(* IEC 61131-3 sources: TetherPLC/compat/tc3 (part 3) *)

(* ---- tc3_mc2_ah.st ---- *)
// Tc3_MC2_AdvancedHoming — user-programmable homing sequences.
//
// All 16 documented APIs over the builtin FB_MotionAxis
// (tplc-motion service), flattened to this dialect:
//
//   AXIS_REF                -> Axis : UDINT (FB_MotionAxis handle)
//   MC_HomingParameter      -> 15 VAR_IN_OUT members P_* (Stored flag
//                             plus the NC soft-limit/lag/vel-diff and
//                             drive torque Stored/Actual fields; the
//                             sim exposes no such drive params so the
//                             fields are pass-through bookkeeping)
//   MC_Ref_Signal_Ref       -> RefLevel : BOOL (the .Level member;
//                             SignalSource/TouchProbe have no sim
//                             equivalent and are dropped)
//   MC_Home_Direction       -> Direction : UDINT
//                             (1=mcPositiveDirection, 3=mcNegative-
//                             Direction, 5=mcSwitchPositive,
//                             7=mcSwitchNegative)
//   MC_Switch_Mode          -> SwitchMode : UDINT
//                             (1=mcOn, 2=mcOff, 3=mcRisingEdge,
//                             4=mcFallingEdge, 5=mcEdgeSwitchPositive,
//                             6=mcEdgeSwitchNegative,
//                             11=mcRisingEdgeInverse,
//                             12=mcFallingEdgeInverse)
//   MC_BufferMode           -> BufferMode : UDINT (not implemented,
//                             accepted and ignored like TwinCAT)
//   ST_Home_Options         -> (empty struct, no member)
//   ST_Home_Options2        -> OptDisableDriveAccess : BOOL
//   ST_Home_Options3        -> OptDisableDriveAccess +
//                             OptInstantLagReduction : BOOL
//   ST_Home_Options4        -> OptDisableDriveAccess +
//                             OptEnableLagErrorDetection : BOOL
//   E_HomingErrorCodes      -> ErrorID values 16#4B90..16#4B98
//
// Motion model: step FBs run a PV-mode (0x6060=3) velocity search at
// Velocity user units/s (0x60FF), poll the OP6 snapshot, and evaluate
// the switch/block condition each scan.  On detection the axis is
// stopped (0x60FF=0), allowed to settle, then the position is assigned
// via a direct 0x6064 write (MC_SetPosition equivalent) unless the FB
// is a "..Detection" variant, which instead returns RecordedPosition.
// The sensor "signal" is the user-fed RefLevel BOOL; the sim has no
// physical switch/encoder inputs.  Block detection uses the
// velocity-undershoot criterion (|VEL_ACTUAL| below
// DetectionVelocityLimit for DetectionVelocityTime); the travel-limit
// clamp added to the velocity modes makes a fixed stop produce that
// undershoot.  TorqueLimit/LagLimit/Acceleration/Deceleration/Jerk are
// accepted but inert (no torque or jerk model in the sim; PV ramps at
// the axis' configured accel/decel).
//
// Internal engine: AH_Run.  Kind codes: 1 absSwitch, 2 absSwitchDet,
// 3 block, 4 blockDet, 5 blockLag, 6 blockLagDet, 7 limitSwitch,
// 8 limitSwitchDet, 9 refPulse, 10 refPulseDet, 11 flyingRefPulse,
// 12 flyingSwitch, 20 distance move (FinishHoming).

// ---- AH_Run: shared homing sequence engine (internal helper) ----
FUNCTION_BLOCK AH_Run
VAR_INPUT
    Execute : BOOL;
    Axis : UDINT;
    Kind : UDINT;
    Direction : UDINT;
    SwitchMode : UDINT;
    RefLevel : BOOL;
    Velocity : LREAL;
    SetPosEn : BOOL;
    SetPosition : LREAL;
    TimeLimit : TIME;
    DistanceLimit : LREAL;
    DetVelLimit : LREAL;
    DetVelTime : TIME;
    LagLimit : LREAL;
    PosLimSw : BOOL;
    NegLimSw : BOOL;
    Distance : LREAL;
    ParamIn : BOOL;
END_VAR
VAR_OUTPUT
    Done : BOOL;
    Busy : BOOL;
    Active : BOOL;
    CommandAborted : BOOL;
    Error : BOOL;
    ErrorID : UDINT;
    RecordedPosition : LREAL;
    ParamOut : BOOL;
END_VAR
VAR
    ax : FB_MotionAxis;
    clk : TON;
    exPrev : BOOL;
    phase : UDINT;          // 0 idle, 1 search, 2 settle, 3 distmove, 4 observe
    refPrev : BOOL;
    moveDir : DINT;
    startPos : DINT;
    startNs : LINT;
    detNs : LINT;           // undershoot start, -1 = not undershooting
    velCmd : DINT;
    pendSet : BOOL;
    recPos : LREAL;
    distGoal : DINT;
    nowNs : LINT;
    pos : DINT;
    vel : DINT;
    cond : BOOL;
    isSwitch : BOOL;
    isBlock : BOOL;
    isDet : BOOL;
    edge : BOOL;
    pStored : BOOL;
END_VAR
    clk(IN := TRUE, PT := T#1000000h);
    ax.AXIS := Axis;
    ax.OP := 3; ax();
    ax.OP := 6; ax();
    Done := FALSE; Busy := FALSE; Active := FALSE;
    CommandAborted := FALSE; Error := FALSE; ErrorID := 0;
    RecordedPosition := 0.0;
    nowNs := TIME_TO_LINT(clk.ET);
    pos := ax.POS_ACTUAL;
    vel := ax.VEL_ACTUAL;
    pStored := ParamIn;
    isSwitch := (Kind >= 1) AND (Kind <= 2) OR (Kind >= 7) AND (Kind <= 10);
    isBlock := (Kind >= 3) AND (Kind <= 6);
    isDet := (Kind = 2) OR (Kind = 4) OR (Kind = 6) OR (Kind = 8)
             OR (Kind = 10);
    edge := Execute AND NOT exPrev;
    exPrev := Execute;

    IF phase = 0 THEN
        IF edge THEN
            // ---- validation ----
            IF Kind <> 11 AND Kind <> 12 AND Velocity <= 0.0 THEN
                Error := TRUE; ErrorID := 16#4B93;   // MC_HOMINGERROR_MODE
            ELSIF Kind <= 12 AND DistanceLimit < 0.0 THEN
                Error := TRUE; ErrorID := 16#4B96;   // DISTANCELIMIT
            ELSIF (Kind >= 1) AND (Kind <= 10)
                  AND Direction <> 1 AND Direction <> 3
                  AND Direction <> 5 AND Direction <> 7 THEN
                Error := TRUE; ErrorID := 16#4B91;   // DIRECTION
            ELSIF isSwitch AND SwitchMode <> 1 AND SwitchMode <> 2
                  AND SwitchMode <> 3 AND SwitchMode <> 4
                  AND SwitchMode <> 5 AND SwitchMode <> 6
                  AND SwitchMode <> 11 AND SwitchMode <> 12 THEN
                Error := TRUE; ErrorID := 16#4B92;   // SWITCHMODE
            ELSE
                // ---- initialise sequence ----
                IF Kind = 20 THEN
                    // distance move (FinishHoming backoff)
                    IF Distance = 0.0 THEN
                        pStored := FALSE;
                        Done := TRUE;
                    ELSE
                        moveDir := 1;
                        IF Distance < 0.0 THEN moveDir := -1; END_IF;
                        startPos := pos; startNs := nowNs; detNs := -1;
                        distGoal := pos + LREAL_TO_DINT(Distance);
                        refPrev := RefLevel;
                        pStored := TRUE;
                        velCmd := LREAL_TO_DINT(DINT_TO_LREAL(moveDir)
                                                * Velocity);
                        ax.OP := 5; ax.INDEX := 16#6060; ax.VALUE := 3; ax();
                        ax.OP := 5; ax.INDEX := 16#60FF;
                        ax.VALUE := velCmd; ax();
                        ax.OP := 5; ax.INDEX := 16#6040;
                        ax.VALUE := 16#000F; ax();
                        IF ax.STATUS = 0 THEN
                            phase := 3; Active := TRUE;
                        ELSE
                            Error := TRUE; ErrorID := ax.ERRID;
                            pStored := FALSE;
                        END_IF;
                    END_IF;
                ELSIF Kind = 11 OR Kind = 12 THEN
                    // passive observation, no motion commanded
                    startPos := pos; startNs := nowNs; detNs := -1;
                    refPrev := RefLevel;
                    pStored := TRUE;
                    phase := 4; Active := TRUE;
                ELSE
                    // search move direction
                    moveDir := 1;
                    IF Direction = 3 THEN moveDir := -1; END_IF;
                    IF Direction = 5 THEN
                        moveDir := 1;
                        IF RefLevel THEN moveDir := -1; END_IF;
                    END_IF;
                    IF Direction = 7 THEN
                        moveDir := -1;
                        IF RefLevel THEN moveDir := 1; END_IF;
                    END_IF;
                    startPos := pos; startNs := nowNs; detNs := -1;
                    refPrev := RefLevel;
                    pStored := TRUE;
                    velCmd := LREAL_TO_DINT(DINT_TO_LREAL(moveDir)
                                            * Velocity);
                    ax.OP := 5; ax.INDEX := 16#6060; ax.VALUE := 3; ax();
                    ax.OP := 5; ax.INDEX := 16#60FF; ax.VALUE := velCmd; ax();
                    ax.OP := 5; ax.INDEX := 16#6040; ax.VALUE := 16#000F; ax();
                    IF ax.STATUS = 0 THEN
                        phase := 1; Active := TRUE;
                    ELSE
                        Error := TRUE; ErrorID := ax.ERRID;
                        pStored := FALSE;
                    END_IF;
                END_IF;
            END_IF;
        END_IF;

    ELSIF phase = 1 THEN
        // ---- search: abort limits then detection ----
        IF (TimeLimit > T#0s) AND
           (nowNs - startNs > TIME_TO_LINT(TimeLimit)) THEN
            ax.OP := 5; ax.INDEX := 16#60FF; ax.VALUE := 0; ax();
            phase := 0; CommandAborted := TRUE;
        ELSIF ABS(DINT_TO_LREAL(pos - startPos)) > DistanceLimit THEN
            ax.OP := 5; ax.INDEX := 16#60FF; ax.VALUE := 0; ax();
            phase := 0; CommandAborted := TRUE;
        ELSIF (PosLimSw AND moveDir > 0) OR (NegLimSw AND moveDir < 0) THEN
            ax.OP := 5; ax.INDEX := 16#60FF; ax.VALUE := 0; ax();
            phase := 0; CommandAborted := TRUE;
        ELSE
            cond := FALSE;
            IF isSwitch THEN
                // MC_Switch_Mode evaluation; inverse variants share
                // the physical edge (approach side is absorbed by
                // the position assignment)
                IF SwitchMode = 1 THEN
                    cond := RefLevel;
                ELSIF SwitchMode = 2 THEN
                    cond := NOT RefLevel;
                ELSIF SwitchMode = 3 OR SwitchMode = 11 THEN
                    cond := RefLevel AND NOT refPrev;
                ELSIF SwitchMode = 4 OR SwitchMode = 12 THEN
                    cond := NOT RefLevel AND refPrev;
                ELSIF SwitchMode = 5 THEN
                    IF moveDir > 0 THEN
                        cond := RefLevel AND NOT refPrev;
                    ELSE
                        cond := NOT RefLevel AND refPrev;
                    END_IF;
                ELSIF SwitchMode = 6 THEN
                    IF moveDir > 0 THEN
                        cond := NOT RefLevel AND refPrev;
                    ELSE
                        cond := RefLevel AND NOT refPrev;
                    END_IF;
                END_IF;
            ELSIF isBlock THEN
                // velocity undershoot below DetVelLimit sustained
                // for DetVelTime; lag-based additionally requires
                // the velocity deficit proxy above LagLimit
                IF ABS(vel) < LREAL_TO_DINT(DetVelLimit) THEN
                    IF detNs < 0 THEN detNs := nowNs; END_IF;
                    IF nowNs - detNs >= TIME_TO_LINT(DetVelTime)
                       AND (Kind < 5 OR
                            ABS(velCmd - vel) > LREAL_TO_DINT(LagLimit)) THEN
                        cond := TRUE;
                    END_IF;
                ELSE
                    detNs := -1;
                END_IF;
            END_IF;
            refPrev := RefLevel;
            IF cond THEN
                ax.OP := 5; ax.INDEX := 16#60FF; ax.VALUE := 0; ax();
                recPos := DINT_TO_LREAL(pos);
                pendSet := SetPosEn AND NOT isDet;
                phase := 2; Active := TRUE;
            ELSE
                Active := TRUE; Busy := TRUE;
            END_IF;
        END_IF;

    ELSIF phase = 2 THEN
        // ---- settle: wait for the velocity ramp-down, then assign
        // the position (or report RecordedPosition) ----
        Active := TRUE; Busy := TRUE;
        IF ABS(vel) <= 1 THEN
            IF pendSet THEN
                ax.OP := 5; ax.INDEX := 16#6064;
                ax.VALUE := LREAL_TO_DINT(SetPosition); ax();
                IF ax.STATUS <> 0 THEN
                    Error := TRUE; ErrorID := ax.ERRID;
                    phase := 0;
                ELSE
                    phase := 0; Done := TRUE;
                    IF Kind = 20 THEN pStored := FALSE; END_IF;
                END_IF;
            ELSE
                IF isDet THEN RecordedPosition := recPos; END_IF;
                phase := 0; Done := TRUE;
                IF Kind = 20 THEN pStored := FALSE; END_IF;
            END_IF;
        END_IF;

    ELSIF phase = 3 THEN
        // ---- distance move: stop at the goal ----
        Active := TRUE; Busy := TRUE;
        IF (moveDir > 0 AND pos >= distGoal)
           OR (moveDir < 0 AND pos <= distGoal) THEN
            ax.OP := 5; ax.INDEX := 16#60FF; ax.VALUE := 0; ax();
            phase := 2;   // reuse settle; pendSet stays FALSE
            pendSet := FALSE;
        END_IF;
        IF (TimeLimit > T#0s) AND
           (nowNs - startNs > TIME_TO_LINT(TimeLimit)) THEN
            ax.OP := 5; ax.INDEX := 16#60FF; ax.VALUE := 0; ax();
            phase := 0; CommandAborted := TRUE; pStored := FALSE;
        END_IF;

    ELSIF phase = 4 THEN
        // ---- passive observation: no motion commanded ----
        Active := TRUE; Busy := TRUE;
        cond := FALSE;
        IF Kind = 11 THEN
            cond := RefLevel AND NOT refPrev;   // encoder zero pulse
        ELSE
            // flying switch: same MC_Switch_Mode evaluation,
            // direction taken as +1 (no search direction)
            IF SwitchMode = 1 THEN cond := RefLevel;
            ELSIF SwitchMode = 2 THEN cond := NOT RefLevel;
            ELSIF SwitchMode = 3 OR SwitchMode = 11 THEN
                cond := RefLevel AND NOT refPrev;
            ELSIF SwitchMode = 4 OR SwitchMode = 12 THEN
                cond := NOT RefLevel AND refPrev;
            ELSIF SwitchMode = 5 THEN
                cond := RefLevel AND NOT refPrev;
            ELSIF SwitchMode = 6 THEN
                cond := NOT RefLevel AND refPrev;
            END_IF;
        END_IF;
        refPrev := RefLevel;
        IF (TimeLimit > T#0s) AND
           (nowNs - startNs > TIME_TO_LINT(TimeLimit)) THEN
            phase := 0; CommandAborted := TRUE; pStored := FALSE;
        ELSIF ABS(DINT_TO_LREAL(pos - startPos)) > DistanceLimit THEN
            phase := 0; CommandAborted := TRUE; pStored := FALSE;
        ELSIF cond THEN
            ax.OP := 5; ax.INDEX := 16#6064;
            ax.VALUE := LREAL_TO_DINT(SetPosition); ax();
            IF ax.STATUS = 0 THEN
                phase := 0; Done := TRUE; pStored := FALSE;
            ELSE
                phase := 0; Error := TRUE; ErrorID := ax.ERRID;
                pStored := FALSE;
            END_IF;
        END_IF;
    END_IF;
    ParamOut := pStored;
END_FUNCTION_BLOCK

// ======================= finalizing FBs =======================

// MC_FinishHoming — completes a homing sequence: optional Distance
// backoff move at Velocity, then restores the stored parameters.
FUNCTION_BLOCK MC_FinishHoming
VAR_INPUT
    Execute : BOOL;
    Distance : LREAL;
    Velocity : LREAL;
    Acceleration : LREAL;
    Deceleration : LREAL;
    Jerk : LREAL;
    BufferMode : UDINT;
    OptDisableDriveAccess : BOOL;
END_VAR
VAR_IN_OUT
    Axis : UDINT;
    P_Stored : BOOL;
    P_NcSMin : BOOL;  P_NcSMax : BOOL;
    P_NcSPosDiff : BOOL;  P_NcSVeloDiff : BOOL;
    P_NcAMin : BOOL;  P_NcAMax : BOOL;
    P_NcAPosDiff : BOOL;  P_NcAVeloDiff : BOOL;
    P_DrvSBip : LREAL;  P_DrvSPos : LREAL;  P_DrvSNeg : LREAL;
    P_DrvABip : LREAL;  P_DrvAPos : LREAL;  P_DrvANeg : LREAL;
END_VAR
VAR_OUTPUT
    Done : BOOL;
    Busy : BOOL;
    CommandAborted : BOOL;
    Error : BOOL;
    ErrorID : UDINT;
END_VAR
VAR
    eng : AH_Run;
END_VAR
    eng.Execute := Execute; eng.Axis := Axis; eng.Kind := 20;
    eng.Direction := 1; eng.SwitchMode := 0; eng.RefLevel := FALSE;
    eng.Velocity := Velocity; eng.SetPosEn := FALSE;
    eng.SetPosition := 0.0;
    eng.TimeLimit := T#0s; eng.DistanceLimit := -1.0;
    eng.DetVelLimit := 0.0; eng.DetVelTime := T#0s; eng.LagLimit := 0.0;
    eng.PosLimSw := FALSE; eng.NegLimSw := FALSE;
    eng.Distance := Distance;
    eng.ParamIn := P_Stored;
    eng();
    P_Stored := eng.ParamOut;
    Done := eng.Done; Busy := eng.Busy;
    CommandAborted := eng.CommandAborted;
    Error := eng.Error; ErrorID := eng.ErrorID;
END_FUNCTION_BLOCK

// MC_HomeDirect — completes homing and assigns the axis position
// directly (no motion).  Axis leaves the homing state.
FUNCTION_BLOCK MC_HomeDirect
VAR_INPUT
    Execute : BOOL;
    SetPosition : LREAL;
    BufferMode : UDINT;
    OptDisableDriveAccess : BOOL;
END_VAR
VAR_IN_OUT
    Axis : UDINT;
    P_Stored : BOOL;
    P_NcSMin : BOOL;  P_NcSMax : BOOL;
    P_NcSPosDiff : BOOL;  P_NcSVeloDiff : BOOL;
    P_NcAMin : BOOL;  P_NcAMax : BOOL;
    P_NcAPosDiff : BOOL;  P_NcAVeloDiff : BOOL;
    P_DrvSBip : LREAL;  P_DrvSPos : LREAL;  P_DrvSNeg : LREAL;
    P_DrvABip : LREAL;  P_DrvAPos : LREAL;  P_DrvANeg : LREAL;
END_VAR
VAR_OUTPUT
    Done : BOOL;
    Busy : BOOL;
    Active : BOOL;
    CommandAborted : BOOL;
    Error : BOOL;
    ErrorID : UDINT;
END_VAR
VAR
    ax : FB_MotionAxis;
    exPrev : BOOL;
END_VAR
    ax.AXIS := Axis;
    Done := FALSE; Busy := FALSE; Active := FALSE;
    CommandAborted := FALSE; Error := FALSE; ErrorID := 0;
    IF Execute AND NOT exPrev THEN
        Active := TRUE;
        ax.OP := 5; ax.INDEX := 16#6064;
        ax.VALUE := LREAL_TO_DINT(SetPosition); ax();
        IF ax.STATUS = 0 THEN
            Done := TRUE; Active := FALSE;
            P_Stored := FALSE;
        ELSE
            Error := TRUE; ErrorID := ax.ERRID;
        END_IF;
    END_IF;
    exPrev := Execute;
END_FUNCTION_BLOCK

// MC_AbortHoming — aborts a homing sequence, stops any search move
// and restores the stored parameters.
FUNCTION_BLOCK MC_AbortHoming
VAR_INPUT
    Execute : BOOL;
    OptDisableDriveAccess : BOOL;
END_VAR
VAR_IN_OUT
    Axis : UDINT;
    P_Stored : BOOL;
    P_NcSMin : BOOL;  P_NcSMax : BOOL;
    P_NcSPosDiff : BOOL;  P_NcSVeloDiff : BOOL;
    P_NcAMin : BOOL;  P_NcAMax : BOOL;
    P_NcAPosDiff : BOOL;  P_NcAVeloDiff : BOOL;
    P_DrvSBip : LREAL;  P_DrvSPos : LREAL;  P_DrvSNeg : LREAL;
    P_DrvABip : LREAL;  P_DrvAPos : LREAL;  P_DrvANeg : LREAL;
END_VAR
VAR_OUTPUT
    Done : BOOL;
    Busy : BOOL;
    CommandAborted : BOOL;
    Error : BOOL;
    ErrorID : UDINT;
END_VAR
VAR
    ax : FB_MotionAxis;
    exPrev : BOOL;
END_VAR
    ax.AXIS := Axis;
    Done := FALSE; Busy := FALSE;
    CommandAborted := FALSE; Error := FALSE; ErrorID := 0;
    IF Execute AND NOT exPrev THEN
        ax.OP := 5; ax.INDEX := 16#60FF; ax.VALUE := 0; ax();
        ax.OP := 5; ax.INDEX := 16#6060; ax.VALUE := 0; ax();
        P_Stored := FALSE;
        Done := (ax.STATUS = 0);
        IF ax.STATUS <> 0 THEN Error := TRUE; ErrorID := ax.ERRID; END_IF;
    END_IF;
    exPrev := Execute;
END_FUNCTION_BLOCK

// ==================== referencing (passive) FBs ====================

// MC_AbortPassiveHoming — aborts passive homing.  The sim keeps no
// NC-side passive state, so this reports Done immediately.
FUNCTION_BLOCK MC_AbortPassiveHoming
VAR_INPUT
    Execute : BOOL;
END_VAR
VAR_IN_OUT
    Axis : UDINT;
END_VAR
VAR_OUTPUT
    Done : BOOL;
    Busy : BOOL;
    Active : BOOL;
    CommandAborted : BOOL;
    Error : BOOL;
    ErrorID : UDINT;
END_VAR
VAR
    exPrev : BOOL;
END_VAR
    Done := FALSE; Busy := FALSE; Active := FALSE;
    CommandAborted := FALSE; Error := FALSE; ErrorID := 0;
    IF Execute AND NOT exPrev THEN
        Done := TRUE;
    END_IF;
    exPrev := Execute;
END_FUNCTION_BLOCK

// MC_StepReferenceFlyingRefPulse — latch the position when the
// encoder zero pulse (RefLevel rising edge) arrives during an
// externally driven move, then assign SetPosition.
FUNCTION_BLOCK MC_StepReferenceFlyingRefPulse
VAR_INPUT
    Execute : BOOL;
    RefLevel : BOOL;
    SetPosition : LREAL;
    TimeLimit : TIME;
    DistanceLimit : LREAL;
    BufferMode : UDINT;
END_VAR
VAR_IN_OUT
    Axis : UDINT;
END_VAR
VAR_OUTPUT
    Done : BOOL;
    Busy : BOOL;
    Active : BOOL;
    CommandAborted : BOOL;
    Error : BOOL;
    ErrorID : UDINT;
END_VAR
VAR
    eng : AH_Run;
END_VAR
    eng.Execute := Execute; eng.Axis := Axis; eng.Kind := 11;
    eng.Direction := 1; eng.SwitchMode := 0; eng.RefLevel := RefLevel;
    eng.Velocity := 0.0; eng.SetPosEn := TRUE;
    eng.SetPosition := SetPosition;
    eng.TimeLimit := TimeLimit; eng.DistanceLimit := DistanceLimit;
    eng.DetVelLimit := 0.0; eng.DetVelTime := T#0s; eng.LagLimit := 0.0;
    eng.PosLimSw := FALSE; eng.NegLimSw := FALSE; eng.Distance := 0.0;
    eng.ParamIn := FALSE;
    eng();
    Done := eng.Done; Busy := eng.Busy; Active := eng.Active;
    CommandAborted := eng.CommandAborted;
    Error := eng.Error; ErrorID := eng.ErrorID;
END_FUNCTION_BLOCK

// MC_StepReferenceFlyingSwitch — same as FlyingRefPulse but the
// trigger is a MC_Switch_Mode condition on RefLevel.
FUNCTION_BLOCK MC_StepReferenceFlyingSwitch
VAR_INPUT
    Execute : BOOL;
    SwitchMode : UDINT;
    RefLevel : BOOL;
    SetPosition : LREAL;
    TimeLimit : TIME;
    DistanceLimit : LREAL;
    BufferMode : UDINT;
END_VAR
VAR_IN_OUT
    Axis : UDINT;
END_VAR
VAR_OUTPUT
    Done : BOOL;
    Busy : BOOL;
    Active : BOOL;
    CommandAborted : BOOL;
    Error : BOOL;
    ErrorID : UDINT;
END_VAR
VAR
    eng : AH_Run;
END_VAR
    eng.Execute := Execute; eng.Axis := Axis; eng.Kind := 12;
    eng.Direction := 1; eng.SwitchMode := SwitchMode;
    eng.RefLevel := RefLevel;
    eng.Velocity := 0.0; eng.SetPosEn := TRUE;
    eng.SetPosition := SetPosition;
    eng.TimeLimit := TimeLimit; eng.DistanceLimit := DistanceLimit;
    eng.DetVelLimit := 0.0; eng.DetVelTime := T#0s; eng.LagLimit := 0.0;
    eng.PosLimSw := FALSE; eng.NegLimSw := FALSE; eng.Distance := 0.0;
    eng.ParamIn := FALSE;
    eng();
    Done := eng.Done; Busy := eng.Busy; Active := eng.Active;
    CommandAborted := eng.CommandAborted;
    Error := eng.Error; ErrorID := eng.ErrorID;
END_FUNCTION_BLOCK

// ========================= step FBs =========================

// MC_StepAbsoluteSwitch — searches for an absolutely positioned external switch
FUNCTION_BLOCK MC_StepAbsoluteSwitch
VAR_INPUT
    Execute : BOOL;
    Direction : UDINT;
    SwitchMode : UDINT;
    RefLevel : BOOL;
    Velocity : LREAL;
    Acceleration : LREAL;
    Deceleration : LREAL;
    Jerk : LREAL;
    SetPosition : LREAL;
    TimeLimit : TIME;
    DistanceLimit : LREAL;
    TorqueLimit : LREAL;
    PositiveLimitSwitch : BOOL;
    NegativeLimitSwitch : BOOL;
    BufferMode : UDINT;
    OptDisableDriveAccess : BOOL;
    OptEnableLagErrorDetection : BOOL;
END_VAR
VAR_IN_OUT
    Axis : UDINT;
    P_Stored : BOOL;
    P_NcSMin : BOOL;  P_NcSMax : BOOL;
    P_NcSPosDiff : BOOL;  P_NcSVeloDiff : BOOL;
    P_NcAMin : BOOL;  P_NcAMax : BOOL;
    P_NcAPosDiff : BOOL;  P_NcAVeloDiff : BOOL;
    P_DrvSBip : LREAL;  P_DrvSPos : LREAL;  P_DrvSNeg : LREAL;
    P_DrvABip : LREAL;  P_DrvAPos : LREAL;  P_DrvANeg : LREAL;
END_VAR
VAR_OUTPUT
    Done : BOOL;
    Busy : BOOL;
    Active : BOOL;
    CommandAborted : BOOL;
    Error : BOOL;
    ErrorID : UDINT;
END_VAR
VAR
    eng : AH_Run;
END_VAR
    eng.Execute := Execute; eng.Axis := Axis;
    eng.Kind := 1;
    eng.Direction := Direction;
    eng.SwitchMode := SwitchMode;
    eng.RefLevel := RefLevel;
    eng.Velocity := Velocity;
    eng.SetPosEn := TRUE;
    eng.SetPosition := SetPosition;
    eng.TimeLimit := TimeLimit;
    eng.DistanceLimit := DistanceLimit;
    eng.DetVelLimit := 0.0;
    eng.DetVelTime := T#0s;
    eng.LagLimit := 0.0;
    eng.PosLimSw := PositiveLimitSwitch;
    eng.NegLimSw := NegativeLimitSwitch;
    eng.Distance := 0.0;
    eng.ParamIn := P_Stored;
    eng();
    P_Stored := eng.ParamOut;
    Done := eng.Done; Busy := eng.Busy; Active := eng.Active;
    CommandAborted := eng.CommandAborted;
    Error := eng.Error; ErrorID := eng.ErrorID;
END_FUNCTION_BLOCK

// MC_StepAbsoluteSwitchDetection — absolute switch search; returns RecordedPosition
FUNCTION_BLOCK MC_StepAbsoluteSwitchDetection
VAR_INPUT
    Execute : BOOL;
    Direction : UDINT;
    SwitchMode : UDINT;
    RefLevel : BOOL;
    Velocity : LREAL;
    Acceleration : LREAL;
    Deceleration : LREAL;
    Jerk : LREAL;
    TimeLimit : TIME;
    DistanceLimit : LREAL;
    TorqueLimit : LREAL;
    PositiveLimitSwitch : BOOL;
    NegativeLimitSwitch : BOOL;
    BufferMode : UDINT;
    OptDisableDriveAccess : BOOL;
    OptEnableLagErrorDetection : BOOL;
END_VAR
VAR_IN_OUT
    Axis : UDINT;
    P_Stored : BOOL;
    P_NcSMin : BOOL;  P_NcSMax : BOOL;
    P_NcSPosDiff : BOOL;  P_NcSVeloDiff : BOOL;
    P_NcAMin : BOOL;  P_NcAMax : BOOL;
    P_NcAPosDiff : BOOL;  P_NcAVeloDiff : BOOL;
    P_DrvSBip : LREAL;  P_DrvSPos : LREAL;  P_DrvSNeg : LREAL;
    P_DrvABip : LREAL;  P_DrvAPos : LREAL;  P_DrvANeg : LREAL;
END_VAR
VAR_OUTPUT
    Done : BOOL;
    Busy : BOOL;
    Active : BOOL;
    CommandAborted : BOOL;
    Error : BOOL;
    ErrorID : UDINT;
    RecordedPosition : LREAL;
END_VAR
VAR
    eng : AH_Run;
END_VAR
    eng.Execute := Execute; eng.Axis := Axis;
    eng.Kind := 2;
    eng.Direction := Direction;
    eng.SwitchMode := SwitchMode;
    eng.RefLevel := RefLevel;
    eng.Velocity := Velocity;
    eng.SetPosEn := FALSE;
    eng.SetPosition := 0.0;
    eng.TimeLimit := TimeLimit;
    eng.DistanceLimit := DistanceLimit;
    eng.DetVelLimit := 0.0;
    eng.DetVelTime := T#0s;
    eng.LagLimit := 0.0;
    eng.PosLimSw := PositiveLimitSwitch;
    eng.NegLimSw := NegativeLimitSwitch;
    eng.Distance := 0.0;
    eng.ParamIn := P_Stored;
    eng();
    P_Stored := eng.ParamOut;
    Done := eng.Done; Busy := eng.Busy; Active := eng.Active;
    CommandAborted := eng.CommandAborted;
    Error := eng.Error; ErrorID := eng.ErrorID;
    RecordedPosition := eng.RecordedPosition;
END_FUNCTION_BLOCK

// MC_StepBlock — search for a mechanical fixed stop (velocity undershoot)
FUNCTION_BLOCK MC_StepBlock
VAR_INPUT
    Execute : BOOL;
    Direction : UDINT;
    Velocity : LREAL;
    Acceleration : LREAL;
    Deceleration : LREAL;
    Jerk : LREAL;
    SetPosition : LREAL;
    DetectionVelocityLimit : LREAL;
    DetectionVelocityTime : TIME;
    TimeLimit : TIME;
    DistanceLimit : LREAL;
    TorqueLimit : LREAL;
    TorqueTolerance : LREAL;
    BufferMode : UDINT;
    OptDisableDriveAccess : BOOL;
    OptInstantLagReduction : BOOL;
END_VAR
VAR_IN_OUT
    Axis : UDINT;
    P_Stored : BOOL;
    P_NcSMin : BOOL;  P_NcSMax : BOOL;
    P_NcSPosDiff : BOOL;  P_NcSVeloDiff : BOOL;
    P_NcAMin : BOOL;  P_NcAMax : BOOL;
    P_NcAPosDiff : BOOL;  P_NcAVeloDiff : BOOL;
    P_DrvSBip : LREAL;  P_DrvSPos : LREAL;  P_DrvSNeg : LREAL;
    P_DrvABip : LREAL;  P_DrvAPos : LREAL;  P_DrvANeg : LREAL;
END_VAR
VAR_OUTPUT
    Done : BOOL;
    Busy : BOOL;
    Active : BOOL;
    CommandAborted : BOOL;
    Error : BOOL;
    ErrorID : UDINT;
END_VAR
VAR
    eng : AH_Run;
END_VAR
    eng.Execute := Execute; eng.Axis := Axis;
    eng.Kind := 3;
    eng.Direction := Direction;
    eng.SwitchMode := 0;
    eng.RefLevel := FALSE;
    eng.Velocity := Velocity;
    eng.SetPosEn := TRUE;
    eng.SetPosition := SetPosition;
    eng.TimeLimit := TimeLimit;
    eng.DistanceLimit := DistanceLimit;
    eng.DetVelLimit := DetectionVelocityLimit;
    eng.DetVelTime := DetectionVelocityTime;
    eng.LagLimit := 0.0;
    eng.PosLimSw := FALSE;
    eng.NegLimSw := FALSE;
    eng.Distance := 0.0;
    eng.ParamIn := P_Stored;
    eng();
    P_Stored := eng.ParamOut;
    Done := eng.Done; Busy := eng.Busy; Active := eng.Active;
    CommandAborted := eng.CommandAborted;
    Error := eng.Error; ErrorID := eng.ErrorID;
END_FUNCTION_BLOCK

// MC_StepBlockDetection — block search; returns RecordedPosition
FUNCTION_BLOCK MC_StepBlockDetection
VAR_INPUT
    Execute : BOOL;
    Direction : UDINT;
    Velocity : LREAL;
    Acceleration : LREAL;
    Deceleration : LREAL;
    Jerk : LREAL;
    DetectionVelocityLimit : LREAL;
    DetectionVelocityTime : TIME;
    TimeLimit : TIME;
    DistanceLimit : LREAL;
    TorqueLimit : LREAL;
    TorqueTolerance : LREAL;
    BufferMode : UDINT;
    OptDisableDriveAccess : BOOL;
    OptInstantLagReduction : BOOL;
END_VAR
VAR_IN_OUT
    Axis : UDINT;
    P_Stored : BOOL;
    P_NcSMin : BOOL;  P_NcSMax : BOOL;
    P_NcSPosDiff : BOOL;  P_NcSVeloDiff : BOOL;
    P_NcAMin : BOOL;  P_NcAMax : BOOL;
    P_NcAPosDiff : BOOL;  P_NcAVeloDiff : BOOL;
    P_DrvSBip : LREAL;  P_DrvSPos : LREAL;  P_DrvSNeg : LREAL;
    P_DrvABip : LREAL;  P_DrvAPos : LREAL;  P_DrvANeg : LREAL;
END_VAR
VAR_OUTPUT
    Done : BOOL;
    Busy : BOOL;
    Active : BOOL;
    CommandAborted : BOOL;
    Error : BOOL;
    ErrorID : UDINT;
    RecordedPosition : LREAL;
END_VAR
VAR
    eng : AH_Run;
END_VAR
    eng.Execute := Execute; eng.Axis := Axis;
    eng.Kind := 4;
    eng.Direction := Direction;
    eng.SwitchMode := 0;
    eng.RefLevel := FALSE;
    eng.Velocity := Velocity;
    eng.SetPosEn := FALSE;
    eng.SetPosition := 0.0;
    eng.TimeLimit := TimeLimit;
    eng.DistanceLimit := DistanceLimit;
    eng.DetVelLimit := DetectionVelocityLimit;
    eng.DetVelTime := DetectionVelocityTime;
    eng.LagLimit := 0.0;
    eng.PosLimSw := FALSE;
    eng.NegLimSw := FALSE;
    eng.Distance := 0.0;
    eng.ParamIn := P_Stored;
    eng();
    P_Stored := eng.ParamOut;
    Done := eng.Done; Busy := eng.Busy; Active := eng.Active;
    CommandAborted := eng.CommandAborted;
    Error := eng.Error; ErrorID := eng.ErrorID;
    RecordedPosition := eng.RecordedPosition;
END_FUNCTION_BLOCK

// MC_StepBlockLagBased — block search with lag-error criterion
FUNCTION_BLOCK MC_StepBlockLagBased
VAR_INPUT
    Execute : BOOL;
    Direction : UDINT;
    Velocity : LREAL;
    Acceleration : LREAL;
    Deceleration : LREAL;
    Jerk : LREAL;
    SetPosition : LREAL;
    DetectionVelocityLimit : LREAL;
    DetectionVelocityTime : TIME;
    TimeLimit : TIME;
    DistanceLimit : LREAL;
    TorqueLimit : LREAL;
    LagLimit : LREAL;
    BufferMode : UDINT;
    OptDisableDriveAccess : BOOL;
    OptInstantLagReduction : BOOL;
END_VAR
VAR_IN_OUT
    Axis : UDINT;
    P_Stored : BOOL;
    P_NcSMin : BOOL;  P_NcSMax : BOOL;
    P_NcSPosDiff : BOOL;  P_NcSVeloDiff : BOOL;
    P_NcAMin : BOOL;  P_NcAMax : BOOL;
    P_NcAPosDiff : BOOL;  P_NcAVeloDiff : BOOL;
    P_DrvSBip : LREAL;  P_DrvSPos : LREAL;  P_DrvSNeg : LREAL;
    P_DrvABip : LREAL;  P_DrvAPos : LREAL;  P_DrvANeg : LREAL;
END_VAR
VAR_OUTPUT
    Done : BOOL;
    Busy : BOOL;
    Active : BOOL;
    CommandAborted : BOOL;
    Error : BOOL;
    ErrorID : UDINT;
END_VAR
VAR
    eng : AH_Run;
END_VAR
    eng.Execute := Execute; eng.Axis := Axis;
    eng.Kind := 5;
    eng.Direction := Direction;
    eng.SwitchMode := 0;
    eng.RefLevel := FALSE;
    eng.Velocity := Velocity;
    eng.SetPosEn := TRUE;
    eng.SetPosition := SetPosition;
    eng.TimeLimit := TimeLimit;
    eng.DistanceLimit := DistanceLimit;
    eng.DetVelLimit := DetectionVelocityLimit;
    eng.DetVelTime := DetectionVelocityTime;
    eng.LagLimit := LagLimit;
    eng.PosLimSw := FALSE;
    eng.NegLimSw := FALSE;
    eng.Distance := 0.0;
    eng.ParamIn := P_Stored;
    eng();
    P_Stored := eng.ParamOut;
    Done := eng.Done; Busy := eng.Busy; Active := eng.Active;
    CommandAborted := eng.CommandAborted;
    Error := eng.Error; ErrorID := eng.ErrorID;
END_FUNCTION_BLOCK

// MC_StepBlockLagBasedDetection — lag-based block search; returns RecordedPosition
FUNCTION_BLOCK MC_StepBlockLagBasedDetection
VAR_INPUT
    Execute : BOOL;
    Direction : UDINT;
    Velocity : LREAL;
    Acceleration : LREAL;
    Deceleration : LREAL;
    Jerk : LREAL;
    SetPosition : LREAL;
    DetectionVelocityLimit : LREAL;
    DetectionVelocityTime : TIME;
    TimeLimit : TIME;
    DistanceLimit : LREAL;
    TorqueLimit : LREAL;
    LagLimit : LREAL;
    BufferMode : UDINT;
    OptDisableDriveAccess : BOOL;
    OptInstantLagReduction : BOOL;
END_VAR
VAR_IN_OUT
    Axis : UDINT;
    P_Stored : BOOL;
    P_NcSMin : BOOL;  P_NcSMax : BOOL;
    P_NcSPosDiff : BOOL;  P_NcSVeloDiff : BOOL;
    P_NcAMin : BOOL;  P_NcAMax : BOOL;
    P_NcAPosDiff : BOOL;  P_NcAVeloDiff : BOOL;
    P_DrvSBip : LREAL;  P_DrvSPos : LREAL;  P_DrvSNeg : LREAL;
    P_DrvABip : LREAL;  P_DrvAPos : LREAL;  P_DrvANeg : LREAL;
END_VAR
VAR_OUTPUT
    Done : BOOL;
    Busy : BOOL;
    Active : BOOL;
    CommandAborted : BOOL;
    Error : BOOL;
    ErrorID : UDINT;
    RecordedPosition : LREAL;
END_VAR
VAR
    eng : AH_Run;
END_VAR
    eng.Execute := Execute; eng.Axis := Axis;
    eng.Kind := 6;
    eng.Direction := Direction;
    eng.SwitchMode := 0;
    eng.RefLevel := FALSE;
    eng.Velocity := Velocity;
    eng.SetPosEn := FALSE;
    eng.SetPosition := 0.0;
    eng.TimeLimit := TimeLimit;
    eng.DistanceLimit := DistanceLimit;
    eng.DetVelLimit := DetectionVelocityLimit;
    eng.DetVelTime := DetectionVelocityTime;
    eng.LagLimit := LagLimit;
    eng.PosLimSw := FALSE;
    eng.NegLimSw := FALSE;
    eng.Distance := 0.0;
    eng.ParamIn := P_Stored;
    eng();
    P_Stored := eng.ParamOut;
    Done := eng.Done; Busy := eng.Busy; Active := eng.Active;
    CommandAborted := eng.CommandAborted;
    Error := eng.Error; ErrorID := eng.ErrorID;
    RecordedPosition := eng.RecordedPosition;
END_FUNCTION_BLOCK

// MC_StepLimitSwitch — search for a hardware limit switch
FUNCTION_BLOCK MC_StepLimitSwitch
VAR_INPUT
    Execute : BOOL;
    Direction : UDINT;
    LimitSwitchMode : UDINT;
    LimitSwitchLevel : BOOL;
    Velocity : LREAL;
    Acceleration : LREAL;
    Deceleration : LREAL;
    Jerk : LREAL;
    SetPosition : LREAL;
    TimeLimit : TIME;
    DistanceLimit : LREAL;
    TorqueLimit : LREAL;
    BufferMode : UDINT;
    OptDisableDriveAccess : BOOL;
    OptEnableLagErrorDetection : BOOL;
END_VAR
VAR_IN_OUT
    Axis : UDINT;
    P_Stored : BOOL;
    P_NcSMin : BOOL;  P_NcSMax : BOOL;
    P_NcSPosDiff : BOOL;  P_NcSVeloDiff : BOOL;
    P_NcAMin : BOOL;  P_NcAMax : BOOL;
    P_NcAPosDiff : BOOL;  P_NcAVeloDiff : BOOL;
    P_DrvSBip : LREAL;  P_DrvSPos : LREAL;  P_DrvSNeg : LREAL;
    P_DrvABip : LREAL;  P_DrvAPos : LREAL;  P_DrvANeg : LREAL;
END_VAR
VAR_OUTPUT
    Done : BOOL;
    Busy : BOOL;
    Active : BOOL;
    CommandAborted : BOOL;
    Error : BOOL;
    ErrorID : UDINT;
END_VAR
VAR
    eng : AH_Run;
END_VAR
    eng.Execute := Execute; eng.Axis := Axis;
    eng.Kind := 7;
    eng.Direction := Direction;
    eng.SwitchMode := LimitSwitchMode;
    eng.RefLevel := LimitSwitchLevel;
    eng.Velocity := Velocity;
    eng.SetPosEn := TRUE;
    eng.SetPosition := SetPosition;
    eng.TimeLimit := TimeLimit;
    eng.DistanceLimit := DistanceLimit;
    eng.DetVelLimit := 0.0;
    eng.DetVelTime := T#0s;
    eng.LagLimit := 0.0;
    eng.PosLimSw := FALSE;
    eng.NegLimSw := FALSE;
    eng.Distance := 0.0;
    eng.ParamIn := P_Stored;
    eng();
    P_Stored := eng.ParamOut;
    Done := eng.Done; Busy := eng.Busy; Active := eng.Active;
    CommandAborted := eng.CommandAborted;
    Error := eng.Error; ErrorID := eng.ErrorID;
END_FUNCTION_BLOCK

// MC_StepLimitSwitchDetection — limit switch search; returns RecordedPosition
FUNCTION_BLOCK MC_StepLimitSwitchDetection
VAR_INPUT
    Execute : BOOL;
    Direction : UDINT;
    LimitSwitchMode : UDINT;
    LimitSwitchLevel : BOOL;
    Velocity : LREAL;
    Acceleration : LREAL;
    Deceleration : LREAL;
    Jerk : LREAL;
    TimeLimit : TIME;
    DistanceLimit : LREAL;
    TorqueLimit : LREAL;
    BufferMode : UDINT;
    OptDisableDriveAccess : BOOL;
    OptEnableLagErrorDetection : BOOL;
END_VAR
VAR_IN_OUT
    Axis : UDINT;
    P_Stored : BOOL;
    P_NcSMin : BOOL;  P_NcSMax : BOOL;
    P_NcSPosDiff : BOOL;  P_NcSVeloDiff : BOOL;
    P_NcAMin : BOOL;  P_NcAMax : BOOL;
    P_NcAPosDiff : BOOL;  P_NcAVeloDiff : BOOL;
    P_DrvSBip : LREAL;  P_DrvSPos : LREAL;  P_DrvSNeg : LREAL;
    P_DrvABip : LREAL;  P_DrvAPos : LREAL;  P_DrvANeg : LREAL;
END_VAR
VAR_OUTPUT
    Done : BOOL;
    Busy : BOOL;
    Active : BOOL;
    CommandAborted : BOOL;
    Error : BOOL;
    ErrorID : UDINT;
    RecordedPosition : LREAL;
END_VAR
VAR
    eng : AH_Run;
END_VAR
    eng.Execute := Execute; eng.Axis := Axis;
    eng.Kind := 8;
    eng.Direction := Direction;
    eng.SwitchMode := LimitSwitchMode;
    eng.RefLevel := LimitSwitchLevel;
    eng.Velocity := Velocity;
    eng.SetPosEn := FALSE;
    eng.SetPosition := 0.0;
    eng.TimeLimit := TimeLimit;
    eng.DistanceLimit := DistanceLimit;
    eng.DetVelLimit := 0.0;
    eng.DetVelTime := T#0s;
    eng.LagLimit := 0.0;
    eng.PosLimSw := FALSE;
    eng.NegLimSw := FALSE;
    eng.Distance := 0.0;
    eng.ParamIn := P_Stored;
    eng();
    P_Stored := eng.ParamOut;
    Done := eng.Done; Busy := eng.Busy; Active := eng.Active;
    CommandAborted := eng.CommandAborted;
    Error := eng.Error; ErrorID := eng.ErrorID;
    RecordedPosition := eng.RecordedPosition;
END_FUNCTION_BLOCK

// MC_StepReferencePulse — search for the encoder zero pulse
FUNCTION_BLOCK MC_StepReferencePulse
VAR_INPUT
    Execute : BOOL;
    Direction : UDINT;
    SwitchMode : UDINT;
    RefLevel : BOOL;
    Velocity : LREAL;
    Acceleration : LREAL;
    Deceleration : LREAL;
    Jerk : LREAL;
    SetPosition : LREAL;
    TimeLimit : TIME;
    DistanceLimit : LREAL;
    TorqueLimit : LREAL;
    BufferMode : UDINT;
    OptDisableDriveAccess : BOOL;
    OptEnableLagErrorDetection : BOOL;
END_VAR
VAR_IN_OUT
    Axis : UDINT;
    P_Stored : BOOL;
    P_NcSMin : BOOL;  P_NcSMax : BOOL;
    P_NcSPosDiff : BOOL;  P_NcSVeloDiff : BOOL;
    P_NcAMin : BOOL;  P_NcAMax : BOOL;
    P_NcAPosDiff : BOOL;  P_NcAVeloDiff : BOOL;
    P_DrvSBip : LREAL;  P_DrvSPos : LREAL;  P_DrvSNeg : LREAL;
    P_DrvABip : LREAL;  P_DrvAPos : LREAL;  P_DrvANeg : LREAL;
END_VAR
VAR_OUTPUT
    Done : BOOL;
    Busy : BOOL;
    Active : BOOL;
    CommandAborted : BOOL;
    Error : BOOL;
    ErrorID : UDINT;
END_VAR
VAR
    eng : AH_Run;
END_VAR
    eng.Execute := Execute; eng.Axis := Axis;
    eng.Kind := 9;
    eng.Direction := Direction;
    eng.SwitchMode := SwitchMode;
    eng.RefLevel := RefLevel;
    eng.Velocity := Velocity;
    eng.SetPosEn := TRUE;
    eng.SetPosition := SetPosition;
    eng.TimeLimit := TimeLimit;
    eng.DistanceLimit := DistanceLimit;
    eng.DetVelLimit := 0.0;
    eng.DetVelTime := T#0s;
    eng.LagLimit := 0.0;
    eng.PosLimSw := FALSE;
    eng.NegLimSw := FALSE;
    eng.Distance := 0.0;
    eng.ParamIn := P_Stored;
    eng();
    P_Stored := eng.ParamOut;
    Done := eng.Done; Busy := eng.Busy; Active := eng.Active;
    CommandAborted := eng.CommandAborted;
    Error := eng.Error; ErrorID := eng.ErrorID;
END_FUNCTION_BLOCK

// MC_StepReferencePulseDetection — zero pulse search; returns RecordedPosition
FUNCTION_BLOCK MC_StepReferencePulseDetection
VAR_INPUT
    Execute : BOOL;
    Direction : UDINT;
    SwitchMode : UDINT;
    RefLevel : BOOL;
    Velocity : LREAL;
    Acceleration : LREAL;
    Deceleration : LREAL;
    Jerk : LREAL;
    TimeLimit : TIME;
    DistanceLimit : LREAL;
    TorqueLimit : LREAL;
    BufferMode : UDINT;
    OptDisableDriveAccess : BOOL;
    OptEnableLagErrorDetection : BOOL;
END_VAR
VAR_IN_OUT
    Axis : UDINT;
    P_Stored : BOOL;
    P_NcSMin : BOOL;  P_NcSMax : BOOL;
    P_NcSPosDiff : BOOL;  P_NcSVeloDiff : BOOL;
    P_NcAMin : BOOL;  P_NcAMax : BOOL;
    P_NcAPosDiff : BOOL;  P_NcAVeloDiff : BOOL;
    P_DrvSBip : LREAL;  P_DrvSPos : LREAL;  P_DrvSNeg : LREAL;
    P_DrvABip : LREAL;  P_DrvAPos : LREAL;  P_DrvANeg : LREAL;
END_VAR
VAR_OUTPUT
    Done : BOOL;
    Busy : BOOL;
    Active : BOOL;
    CommandAborted : BOOL;
    Error : BOOL;
    ErrorID : UDINT;
    RecordedPosition : LREAL;
END_VAR
VAR
    eng : AH_Run;
END_VAR
    eng.Execute := Execute; eng.Axis := Axis;
    eng.Kind := 10;
    eng.Direction := Direction;
    eng.SwitchMode := SwitchMode;
    eng.RefLevel := RefLevel;
    eng.Velocity := Velocity;
    eng.SetPosEn := FALSE;
    eng.SetPosition := 0.0;
    eng.TimeLimit := TimeLimit;
    eng.DistanceLimit := DistanceLimit;
    eng.DetVelLimit := 0.0;
    eng.DetVelTime := T#0s;
    eng.LagLimit := 0.0;
    eng.PosLimSw := FALSE;
    eng.NegLimSw := FALSE;
    eng.Distance := 0.0;
    eng.ParamIn := P_Stored;
    eng();
    P_Stored := eng.ParamOut;
    Done := eng.Done; Busy := eng.Busy; Active := eng.Active;
    CommandAborted := eng.CommandAborted;
    Error := eng.Error; ErrorID := eng.ErrorID;
    RecordedPosition := eng.RecordedPosition;
END_FUNCTION_BLOCK

(* ---- tc3_mc3cam.st ---- *)
// Tc3_Mc3Camming — MC3 phasing and gear-in-position blocks
// (TF55xx_MC3 camming/phasing subset).
//
// Implemented PLC-side over FB_MotionAxis, mirroring the MC_GearIn
// feedforward pattern in tc2_mc2.st: while the command is active
// each scan reads master position (0x6064) and velocity (0x606C),
// computes the slave position target and commands slave velocity
// (PV mode, 0x60FF)
//     velCmd = masterVel + Kp * (target - slavePos)
// The proportional term is the phase correction; Kp = 10 gives a
// ~100 ms position time constant in the simulated drive. Done /
// InSync report once the position error stays inside TOL for
// SUS scans. This is a documented approximation: real phasing and
// gear-in run inside the NC kernel with profile supervision and a
// persistent cam coupling; here the command ends at Done and the
// slave keeps its last velocity command until another motion
// command (MC_HaltPhasing, MC_GearOut, MC_Stop, ...) takes over.
//
//   MC_PhasingAbsolute  target = masterPos + PhaseShift
//   MC_PhasingRelative  target = masterPos + offset0 + PhaseShift
//                      (offset0 = slavePos - masterPos at engage)
//   MC_GearInPos        target = slavePos0 + ratio*(masterPos - masterPos0)
//   MC_HaltPhasing      ramp slave to rest, Done at VEL_ACTUAL = 0
//
// The cam-table FBs (MC_CamIn/Add/Exchange/Remove/Scaling/
// TableSelect/ReadCamInfo) need the NCI path kernel and remain
// deferred; MC_Cam* table storage is covered by tc3_nccam's
// single-table coupling engine, not this API surface.

// convergence window and sustain count shared by all phasing FBs
// (ST has no constants; literals inlined per FB)

FUNCTION_BLOCK MC_PhasingAbsolute
VAR_INPUT
    Execute : BOOL;
    PhaseShift : DINT;
    Velocity : DINT;
    Acceleration : DINT;
    Deceleration : DINT;
    Jerk : DINT;
    Master : UDINT;
    Slave : UDINT;
END_VAR
VAR_OUTPUT
    Done : BOOL;
    Busy : BOOL;
    Error : BOOL;
    ErrorID : UDINT;
END_VAR
VAR
    axM : FB_MotionAxis;
    axS : FB_MotionAxis;
    exPrev : BOOL;
    exEdge : BOOL;
    active : BOOL;
    good : INT;
    mpos : DINT;
    mvel : DINT;
    spos : DINT;
    tgt : DINT;
    vcmd : DINT;
END_VAR
    axM.AXIS := Master;
    axS.AXIS := Slave;
    axM.OP := 3; axM();
    exEdge := Execute AND NOT exPrev; exPrev := Execute;
    Done := FALSE; Error := FALSE; ErrorID := 0;
    IF exEdge AND NOT active THEN
        axS.OP := 5; axS.INDEX := 16#6040; axS.VALUE := 16#000F; axS();
        axS.OP := 5; axS.INDEX := 16#6060; axS.VALUE := 3; axS();
        active := TRUE; good := 0;
    END_IF;
    IF active THEN
        axM.OP := 4; axM.INDEX := 16#6064; axM(); mpos := axM.VALUE;
        axM.OP := 4; axM.INDEX := 16#606C; axM(); mvel := axM.VALUE;
        axS.OP := 4; axS.INDEX := 16#6064; axS(); spos := axS.VALUE;
        tgt := mpos + PhaseShift;
        vcmd := mvel + (tgt - spos) * 10;
        axS.OP := 5; axS.INDEX := 16#60FF; axS.VALUE := vcmd; axS();
        axS.OP := 6; axS();
        IF axS.STATUS < 0 THEN
            Error := TRUE; ErrorID := axS.ERRID; active := FALSE;
        ELSIF ABS(spos - tgt) <= 250 THEN
            good := good + 1;
            IF good >= 5 THEN
                Done := TRUE; active := FALSE;
            END_IF;
        ELSE
            good := 0;
        END_IF;
    END_IF;
    Busy := active;
END_FUNCTION_BLOCK

FUNCTION_BLOCK MC_PhasingRelative
VAR_INPUT
    Execute : BOOL;
    PhaseShift : DINT;
    Velocity : DINT;
    Acceleration : DINT;
    Deceleration : DINT;
    Jerk : DINT;
    Master : UDINT;
    Slave : UDINT;
END_VAR
VAR_OUTPUT
    Done : BOOL;
    Busy : BOOL;
    Error : BOOL;
    ErrorID : UDINT;
END_VAR
VAR
    axM : FB_MotionAxis;
    axS : FB_MotionAxis;
    exPrev : BOOL;
    exEdge : BOOL;
    active : BOOL;
    haveOff : BOOL;
    good : INT;
    off : DINT;
    mpos : DINT;
    mvel : DINT;
    spos : DINT;
    tgt : DINT;
    vcmd : DINT;
END_VAR
    axM.AXIS := Master;
    axS.AXIS := Slave;
    axM.OP := 3; axM();
    exEdge := Execute AND NOT exPrev; exPrev := Execute;
    Done := FALSE; Error := FALSE; ErrorID := 0;
    IF exEdge AND NOT active THEN
        axS.OP := 5; axS.INDEX := 16#6040; axS.VALUE := 16#000F; axS();
        axS.OP := 5; axS.INDEX := 16#6060; axS.VALUE := 3; axS();
        active := TRUE; good := 0; haveOff := FALSE;
    END_IF;
    IF active THEN
        axM.OP := 4; axM.INDEX := 16#6064; axM(); mpos := axM.VALUE;
        axM.OP := 4; axM.INDEX := 16#606C; axM(); mvel := axM.VALUE;
        axS.OP := 4; axS.INDEX := 16#6064; axS(); spos := axS.VALUE;
        IF NOT haveOff THEN
            off := spos - mpos;
            haveOff := TRUE;
        END_IF;
        tgt := mpos + off + PhaseShift;
        vcmd := mvel + (tgt - spos) * 10;
        axS.OP := 5; axS.INDEX := 16#60FF; axS.VALUE := vcmd; axS();
        axS.OP := 6; axS();
        IF axS.STATUS < 0 THEN
            Error := TRUE; ErrorID := axS.ERRID; active := FALSE;
        ELSIF ABS(spos - tgt) <= 250 THEN
            good := good + 1;
            IF good >= 5 THEN
                Done := TRUE; active := FALSE;
            END_IF;
        ELSE
            good := 0;
        END_IF;
    END_IF;
    Busy := active;
END_FUNCTION_BLOCK

FUNCTION_BLOCK MC_GearInPos
VAR_INPUT
    Execute : BOOL;
    RatioNumerator : DINT;
    RatioDenominator : DINT;
    Velocity : DINT;
    Acceleration : DINT;
    Deceleration : DINT;
    Jerk : DINT;
    Master : UDINT;
    Slave : UDINT;
END_VAR
VAR_OUTPUT
    InSync : BOOL;
    Busy : BOOL;
    Error : BOOL;
    ErrorID : UDINT;
END_VAR
VAR
    axM : FB_MotionAxis;
    axS : FB_MotionAxis;
    exPrev : BOOL;
    exEdge : BOOL;
    active : BOOL;
    haveAnchor : BOOL;
    good : INT;
    mpos0 : DINT;
    spos0 : DINT;
    mpos : DINT;
    mvel : DINT;
    spos : DINT;
    tgt : DINT;
    vcmd : DINT;
END_VAR
    axM.AXIS := Master;
    axS.AXIS := Slave;
    axM.OP := 3; axM();
    exEdge := Execute AND NOT exPrev; exPrev := Execute;
    InSync := FALSE; Error := FALSE; ErrorID := 0;
    IF exEdge AND NOT active THEN
        IF RatioDenominator = 0 THEN
            Error := TRUE; ErrorID := 1;
        ELSE
            axS.OP := 5; axS.INDEX := 16#6040; axS.VALUE := 16#000F; axS();
            axS.OP := 5; axS.INDEX := 16#6060; axS.VALUE := 3; axS();
            active := TRUE; good := 0; haveAnchor := FALSE;
        END_IF;
    END_IF;
    IF active THEN
        axM.OP := 4; axM.INDEX := 16#6064; axM(); mpos := axM.VALUE;
        axM.OP := 4; axM.INDEX := 16#606C; axM(); mvel := axM.VALUE;
        axS.OP := 4; axS.INDEX := 16#6064; axS(); spos := axS.VALUE;
        IF NOT haveAnchor THEN
            mpos0 := mpos; spos0 := spos; haveAnchor := TRUE;
        END_IF;
        tgt := spos0 + (mpos - mpos0) * RatioNumerator / RatioDenominator;
        vcmd := mvel * RatioNumerator / RatioDenominator
                + (tgt - spos) * 10;
        axS.OP := 5; axS.INDEX := 16#60FF; axS.VALUE := vcmd; axS();
        axS.OP := 6; axS();
        IF axS.STATUS < 0 THEN
            Error := TRUE; ErrorID := axS.ERRID; active := FALSE;
        ELSIF ABS(spos - tgt) <= 250 THEN
            good := good + 1;
            IF good >= 5 THEN
                InSync := TRUE; active := FALSE;
            END_IF;
        ELSE
            good := 0;
        END_IF;
    END_IF;
    Busy := active;
END_FUNCTION_BLOCK

// ---- MC_HaltPhasing: ramp the slave to rest and disengage ----
FUNCTION_BLOCK MC_HaltPhasing
VAR_INPUT
    Execute : BOOL;
    Deceleration : DINT;
    Jerk : DINT;
    Master : UDINT;
    Slave : UDINT;
END_VAR
VAR_OUTPUT
    Done : BOOL;
    Busy : BOOL;
    Error : BOOL;
    ErrorID : UDINT;
END_VAR
VAR
    axS : FB_MotionAxis;
    exPrev : BOOL;
    exEdge : BOOL;
    active : BOOL;
END_VAR
    axS.AXIS := Slave;
    axS.OP := 3; axS();
    exEdge := Execute AND NOT exPrev; exPrev := Execute;
    Done := FALSE; Error := FALSE; ErrorID := 0;
    IF exEdge AND NOT active THEN
        axS.OP := 5; axS.INDEX := 16#60FF; axS.VALUE := 0; axS();
        active := TRUE;
    END_IF;
    IF active THEN
        axS.OP := 6; axS();
        IF axS.STATUS < 0 THEN
            Error := TRUE; ErrorID := axS.ERRID; active := FALSE;
        ELSIF axS.VEL_ACTUAL = 0 THEN
            Done := TRUE; active := FALSE;
        END_IF;
    END_IF;
    Busy := active;
END_FUNCTION_BLOCK

// ===========================================================================
// Cam table objects + cam coupling FBs (Tc3_Mc3Camming §5.4.3).
//
// TwinCAT models cam tables as MC_CamObject / Type_CouplingFunction1D
// objects with METHOD-based point access; this dialect has no object
// references or METHODs, so a cam object flattens to a UDINT handle in
// the tplc-cam service. FB_CamTable is the compat-side object holder
// (create/write/config edges — the flattened METHOD surface);
// MC_CamTableSelect applies periodic/continuity to a handle;
// MC_CamIn/Add/Exchange bind a slave axis to master+cam and stream the
// interpolated position target over 0x607A (CSP) while the binding
// lives; MC_CamRemove/MC_CamScaling/MC_ReadCamInfo operate on the
// shared binding registry.
//
// Documented deviations: one binding per slave (multi-plate cam
// summation deferred — cam_bind returns E_BOUND), cam tables are
// point lists in axis user units (LREAL storage, DINT boundary like
// tc3_nccam), continuity requirement is stored but not enforced,
// ActivationOptions/BufferMode inputs accepted but not modeled.
// ===========================================================================

// ---- FB_CamTable: flattened MC_CamObject (table holder) ----
FUNCTION_BLOCK FB_CamTable
VAR_INPUT
    WritePt : BOOL;
    PtIndex : UDINT;
    PtMaster : LREAL;
    PtSlave : LREAL;
    ClearTable : BOOL;
    Config : BOOL;
    TableCount : UDINT;
    Periodic : BOOL;
    Continuity : UDINT;
END_VAR
VAR_OUTPUT
    Error : BOOL;
    ErrorID : UDINT;
END_VAR
VAR
    cam : FB_Cam;
    prevWr : BOOL;
    prevClr : BOOL;
    prevCfg : BOOL;
    flags : UDINT;
    Handle : UDINT;   // public: cam object handle for MC_CAM_REF flattening
END_VAR
    Error := FALSE; ErrorID := 0;
    IF Handle = 0 THEN
        cam.OP := 0; cam();
        IF cam.STATUS = 0 THEN Handle := cam.HANDLE; END_IF;
    END_IF;
    IF Handle <> 0 THEN
        cam.HANDLE := Handle;
        IF WritePt AND NOT prevWr THEN
            cam.OP := 2; cam.AUX := PtIndex;
            cam.F1 := PtMaster; cam.F2 := PtSlave; cam();
            IF cam.STATUS <> 0 THEN
                Error := TRUE; ErrorID := cam.ERRID;
            END_IF;
        END_IF;
        IF ClearTable AND NOT prevClr THEN
            cam.OP := 1; cam();
            IF cam.STATUS <> 0 THEN
                Error := TRUE; ErrorID := cam.ERRID;
            END_IF;
        END_IF;
        IF Config AND NOT prevCfg THEN
            flags := Continuity * 2;
            IF Periodic THEN flags := flags + 1; END_IF;
            cam.OP := 3; cam.AUX := TableCount; cam.FLAGS := flags;
            cam();
            IF cam.STATUS <> 0 THEN
                Error := TRUE; ErrorID := cam.ERRID;
            END_IF;
        END_IF;
    END_IF;
    prevWr := WritePt; prevClr := ClearTable; prevCfg := Config;
END_FUNCTION_BLOCK

// shared cam-stream loop shape (inlined per FB; the dialect has no
// inheritance):
//   OP7 bound query -> cam/master/scalings (fresh each scan so
//     MC_CamScaling updates propagate and MC_CamRemove stops the
//     stream when the binding disappears)
//   master POS_ACTUAL -> mt = act*mscale+moff -> OP4 eval -> st
//   st = st*sscale+soff -> write slave 0x607A = LREAL_TO_DINT(st)
//   (CSP position-target streaming, same as tc3_nccam)
//   InSync when |slavePosActual - tgt| <= 250 for 5 scans

FUNCTION_BLOCK MC_CamIn
VAR_INPUT
    Execute : BOOL;
    Master : UDINT;
    Slave : UDINT;
    CamObject : UDINT;
    MasterScaling : LREAL := 1.0;
    MasterOffset : LREAL := 0.0;
    SlaveScaling : LREAL := 1.0;
    SlaveOffset : LREAL := 0.0;
    ActivationMode : UDINT := 0;
    ActivationPosition : LREAL := 0.0;
    ActivationReference : UDINT := 0;
    BufferMode : UDINT := 0;
END_VAR
VAR_OUTPUT
    InSync : BOOL;
    Busy : BOOL;
    Error : BOOL;
    ErrorID : UDINT;
END_VAR
VAR
    cam : FB_Cam;
    axM : FB_MotionAxis;
    axS : FB_MotionAxis;
    exPrev : BOOL;
    exEdge : BOOL;
    good : INT;
    bCam : UDINT;
    bMaster : UDINT;
    mAct : DINT;
    sAct : DINT;
    mt : LREAL;
    st : LREAL;
    tgt : DINT;
    msc : LREAL;
    mofs : LREAL;
    ssc : LREAL;
    sofs : LREAL;
END_VAR
    cam.AUX := Slave;
    cam.OP := 7; cam();
    bCam := cam.HANDLE;
    msc := cam.F1; mofs := cam.F2; ssc := cam.F3; sofs := cam.F4;
    exEdge := Execute AND NOT exPrev; exPrev := Execute;
    InSync := FALSE; Busy := FALSE;
    Error := FALSE; ErrorID := 0;
    IF exEdge THEN
        cam.OP := 6;
        cam.AUX := Slave; cam.AUX2 := Master; cam.HANDLE := CamObject;
        cam.F1 := MasterScaling; cam.F2 := MasterOffset;
        cam.F3 := SlaveScaling; cam.F4 := SlaveOffset;
        cam();
        IF cam.STATUS <> 0 THEN
            Error := TRUE; ErrorID := cam.ERRID;
        END_IF;
    END_IF;
    IF bCam <> 0 AND CamObject <> 0 AND bCam = CamObject THEN
        Busy := TRUE;
        axM.AXIS := bMaster; axM.OP := 3; axM();
        axM.OP := 6; axM(); mAct := axM.POS_ACTUAL;
        mt := DINT_TO_LREAL(mAct) * msc + mofs;
        cam.OP := 4; cam.HANDLE := bCam; cam.F1 := mt; cam();
        st := cam.F2 * ssc + sofs;
        tgt := LREAL_TO_DINT(st);
        axS.AXIS := Slave; axS.OP := 3; axS();
        axS.OP := 6; axS(); sAct := axS.POS_ACTUAL;
        axS.OP := 5; axS.INDEX := 16#607A; axS.VALUE := tgt; axS();
        IF axS.STATUS < 0 THEN
            Error := TRUE; ErrorID := axS.ERRID; Busy := FALSE;
        ELSIF ABS(sAct - tgt) <= 250 THEN
            good := good + 1;
            IF good >= 5 THEN InSync := TRUE; END_IF;
        ELSE
            good := 0;
        END_IF;
    END_IF;
END_FUNCTION_BLOCK

// ---- MC_CamAdd: additional cam coupling (single-binding rule) ----
// Multi-plate summation needs the NC kernel; cam_bind rejects a
// second binding on the same slave, so this behaves like MC_CamIn
// when the slave is free and errors when it is already coupled.
FUNCTION_BLOCK MC_CamAdd
VAR_INPUT
    Execute : BOOL;
    Master : UDINT;
    Slave : UDINT;
    CamObject : UDINT;
    MasterScaling : LREAL := 1.0;
    MasterOffset : LREAL := 0.0;
    SlaveScaling : LREAL := 1.0;
    SlaveOffset : LREAL := 0.0;
    ActivationMode : UDINT := 0;
    ActivationPosition : LREAL := 0.0;
    ActivationReference : UDINT := 0;
    BufferMode : UDINT := 0;
END_VAR
VAR_OUTPUT
    InSync : BOOL;
    Busy : BOOL;
    Error : BOOL;
    ErrorID : UDINT;
END_VAR
VAR
    cam : FB_Cam;
    axM : FB_MotionAxis;
    axS : FB_MotionAxis;
    exPrev : BOOL;
    exEdge : BOOL;
    good : INT;
    bCam : UDINT;
    mAct : DINT;
    sAct : DINT;
    mt : LREAL;
    st : LREAL;
    tgt : DINT;
    msc : LREAL;
    mofs : LREAL;
    ssc : LREAL;
    sofs : LREAL;
END_VAR
    cam.AUX := Slave;
    cam.OP := 7; cam();
    bCam := cam.HANDLE;
    msc := cam.F1; mofs := cam.F2; ssc := cam.F3; sofs := cam.F4;
    exEdge := Execute AND NOT exPrev; exPrev := Execute;
    InSync := FALSE; Busy := FALSE;
    Error := FALSE; ErrorID := 0;
    IF exEdge THEN
        cam.OP := 6;
        cam.AUX := Slave; cam.AUX2 := Master; cam.HANDLE := CamObject;
        cam.F1 := MasterScaling; cam.F2 := MasterOffset;
        cam.F3 := SlaveScaling; cam.F4 := SlaveOffset;
        cam();
        IF cam.STATUS <> 0 THEN
            Error := TRUE; ErrorID := cam.ERRID;
        END_IF;
    END_IF;
    IF bCam <> 0 AND CamObject <> 0 AND bCam = CamObject THEN
        Busy := TRUE;
        axM.AXIS := Master; axM.OP := 3; axM();
        axM.OP := 6; axM(); mAct := axM.POS_ACTUAL;
        mt := DINT_TO_LREAL(mAct) * msc + mofs;
        cam.OP := 4; cam.HANDLE := bCam; cam.F1 := mt; cam();
        st := cam.F2 * ssc + sofs;
        tgt := LREAL_TO_DINT(st);
        axS.AXIS := Slave; axS.OP := 3; axS();
        axS.OP := 6; axS(); sAct := axS.POS_ACTUAL;
        axS.OP := 5; axS.INDEX := 16#607A; axS.VALUE := tgt; axS();
        IF axS.STATUS < 0 THEN
            Error := TRUE; ErrorID := axS.ERRID; Busy := FALSE;
        ELSIF ABS(sAct - tgt) <= 250 THEN
            good := good + 1;
            IF good >= 5 THEN InSync := TRUE; END_IF;
        ELSE
            good := 0;
        END_IF;
    END_IF;
END_FUNCTION_BLOCK

// ---- MC_CamExchange: swap the slave's cam coupling ----
FUNCTION_BLOCK MC_CamExchange
VAR_INPUT
    Execute : BOOL;
    Master : UDINT;
    Slave : UDINT;
    CamObjectToRemove : UDINT;
    CamObjectToAdd : UDINT;
    MasterScaling : LREAL := 1.0;
    MasterOffset : LREAL := 0.0;
    SlaveScaling : LREAL := 1.0;
    SlaveOffset : LREAL := 0.0;
    ActivationMode : UDINT := 0;
    ActivationPosition : LREAL := 0.0;
    ActivationReference : UDINT := 0;
    BufferMode : UDINT := 0;
END_VAR
VAR_OUTPUT
    InSync : BOOL;
    Busy : BOOL;
    Error : BOOL;
    ErrorID : UDINT;
END_VAR
VAR
    cam : FB_Cam;
    axM : FB_MotionAxis;
    axS : FB_MotionAxis;
    exPrev : BOOL;
    exEdge : BOOL;
    good : INT;
    myCam : UDINT;
    mAct : DINT;
    sAct : DINT;
    mt : LREAL;
    st : LREAL;
    tgt : DINT;
    msc : LREAL;
    mofs : LREAL;
    ssc : LREAL;
    sofs : LREAL;
END_VAR
    cam.AUX := Slave;
    cam.OP := 7; cam();
    msc := cam.F1; mofs := cam.F2; ssc := cam.F3; sofs := cam.F4;
    exEdge := Execute AND NOT exPrev; exPrev := Execute;
    InSync := FALSE; Busy := FALSE;
    Error := FALSE; ErrorID := 0;
    IF exEdge THEN
        // remove must target the currently bound cam object
        cam.OP := 8; cam.AUX := Slave; cam.HANDLE := CamObjectToRemove;
        cam();
        IF cam.STATUS = 0 THEN
            cam.OP := 6;
            cam.AUX := Slave; cam.AUX2 := Master;
            cam.HANDLE := CamObjectToAdd;
            cam.F1 := MasterScaling; cam.F2 := MasterOffset;
            cam.F3 := SlaveScaling; cam.F4 := SlaveOffset;
            cam();
            IF cam.STATUS = 0 THEN myCam := CamObjectToAdd; END_IF;
        END_IF;
        IF cam.STATUS <> 0 THEN
            Error := TRUE; ErrorID := cam.ERRID;
        END_IF;
    END_IF;
    IF myCam <> 0 THEN
        Busy := TRUE;
        axM.AXIS := Master; axM.OP := 3; axM();
        axM.OP := 6; axM(); mAct := axM.POS_ACTUAL;
        mt := DINT_TO_LREAL(mAct) * msc + mofs;
        cam.OP := 4; cam.HANDLE := myCam; cam.F1 := mt; cam();
        st := cam.F2 * ssc + sofs;
        tgt := LREAL_TO_DINT(st);
        axS.AXIS := Slave; axS.OP := 3; axS();
        axS.OP := 6; axS(); sAct := axS.POS_ACTUAL;
        axS.OP := 5; axS.INDEX := 16#607A; axS.VALUE := tgt; axS();
        IF axS.STATUS < 0 THEN
            Error := TRUE; ErrorID := axS.ERRID; Busy := FALSE;
        ELSIF ABS(sAct - tgt) <= 250 THEN
            good := good + 1;
            IF good >= 5 THEN InSync := TRUE; END_IF;
        ELSE
            good := 0;
        END_IF;
    END_IF;
END_FUNCTION_BLOCK

// ---- MC_CamRemove: drop the slave's cam coupling ----
FUNCTION_BLOCK MC_CamRemove
VAR_INPUT
    Execute : BOOL;
    Slave : UDINT;
    CamObject : UDINT;
    ActivationMode : UDINT := 0;
    ActivationPosition : LREAL := 0.0;
    ActivationReference : UDINT := 0;
END_VAR
VAR_OUTPUT
    Done : BOOL;
    Busy : BOOL;
    Error : BOOL;
    ErrorID : UDINT;
END_VAR
VAR
    cam : FB_Cam;
    exPrev : BOOL;
    exEdge : BOOL;
END_VAR
    cam.AUX := Slave;
    cam.OP := 7; cam();
    exEdge := Execute AND NOT exPrev; exPrev := Execute;
    Done := FALSE; Busy := FALSE;
    Error := FALSE; ErrorID := 0;
    IF exEdge THEN
        cam.OP := 8; cam.AUX := Slave; cam.HANDLE := CamObject; cam();
        IF cam.STATUS = 0 THEN
            Done := TRUE;
        ELSE
            Error := TRUE; ErrorID := cam.ERRID;
        END_IF;
    END_IF;
END_FUNCTION_BLOCK

// ---- MC_CamScaling: update coupling scalings on a bound slave ----
FUNCTION_BLOCK MC_CamScaling
VAR_INPUT
    Execute : BOOL;
    Slave : UDINT;
    CamObject : UDINT;
    MasterScaling : LREAL := 1.0;
    MasterOffset : LREAL := 0.0;
    SlaveScaling : LREAL := 1.0;
    SlaveOffset : LREAL := 0.0;
    ActivationMode : UDINT := 0;
    ActivationPosition : LREAL := 0.0;
    ActivationReference : UDINT := 0;
END_VAR
VAR_OUTPUT
    Done : BOOL;
    Busy : BOOL;
    Error : BOOL;
    ErrorID : UDINT;
END_VAR
VAR
    cam : FB_Cam;
    exPrev : BOOL;
    exEdge : BOOL;
END_VAR
    cam.AUX := Slave;
    exEdge := Execute AND NOT exPrev; exPrev := Execute;
    Done := FALSE; Busy := FALSE;
    Error := FALSE; ErrorID := 0;
    IF exEdge THEN
        cam.OP := 9;
        cam.AUX := Slave;
        cam.F1 := MasterScaling; cam.F2 := MasterOffset;
        cam.F3 := SlaveScaling; cam.F4 := SlaveOffset;
        cam();
        IF cam.STATUS = 0 THEN
            Done := TRUE;
        ELSE
            Error := TRUE; ErrorID := cam.ERRID;
        END_IF;
    END_IF;
END_FUNCTION_BLOCK

// ---- MC_CamTableSelect: apply periodic/continuity to a cam object ----
// CamRef and CamObject both flatten to the same UDINT handle (the
// object IS the table); CamObjectOut echoes the configured handle.
FUNCTION_BLOCK MC_CamTableSelect
VAR_INPUT
    Execute : BOOL;
    CamRef : UDINT;
    Periodic : BOOL;
    ContinuityRequirement : UDINT := 0;
    CamObjectIn : UDINT := 0;
END_VAR
VAR_OUTPUT
    CamObjectOut : UDINT;
    Done : BOOL;
    Busy : BOOL;
    Error : BOOL;
    ErrorID : UDINT;
END_VAR
VAR
    cam : FB_Cam;
    exPrev : BOOL;
    exEdge : BOOL;
    flags : UDINT;
    h : UDINT;
END_VAR
    h := CamObjectIn;
    IF h = 0 THEN h := CamRef; END_IF;
    exEdge := Execute AND NOT exPrev; exPrev := Execute;
    CamObjectOut := h;
    Done := FALSE; Busy := FALSE;
    Error := FALSE; ErrorID := 0;
    IF exEdge AND h <> 0 THEN
        flags := ContinuityRequirement * 2;
        IF Periodic THEN flags := flags + 1; END_IF;
        cam.OP := 3; cam.HANDLE := h; cam.AUX := 0; cam.FLAGS := flags;
        cam();
        IF cam.STATUS = 0 THEN
            Done := TRUE;
        ELSE
            Error := TRUE; ErrorID := cam.ERRID;
        END_IF;
    END_IF;
END_FUNCTION_BLOCK

// ---- MC_ReadCamInfo: report the slave's cam coupling ----
// CouplingInfo[] flattens to scalar outputs for the (single)
// binding: CamHandle/MasterAxis/InSync/SlaveScaling.
FUNCTION_BLOCK MC_ReadCamInfo
VAR_INPUT
    Execute : BOOL;
    Slave : UDINT;
    NumberOfCouplings : UDINT := 8;
END_VAR
VAR_OUTPUT
    Done : BOOL;
    Busy : BOOL;
    Error : BOOL;
    ErrorID : UDINT;
    NumberOfCouplingsFound : UDINT;
    CamHandle : UDINT;
    MasterAxis : UDINT;
    CouplingInSync : BOOL;
    SlaveScaling : LREAL;
END_VAR
VAR
    cam : FB_Cam;
    exPrev : BOOL;
    exEdge : BOOL;
END_VAR
    cam.AUX := Slave;
    cam.OP := 7; cam();
    exEdge := Execute AND NOT exPrev; exPrev := Execute;
    Done := FALSE; Busy := FALSE;
    Error := FALSE; ErrorID := 0;
    NumberOfCouplingsFound := 0;
    CamHandle := 0; MasterAxis := 0;
    CouplingInSync := FALSE; SlaveScaling := 1.0;
    IF exEdge THEN
        IF cam.STATUS = 0 THEN
            Done := TRUE;
            IF cam.HANDLE <> 0 THEN
                NumberOfCouplingsFound := 1;
                CamHandle := cam.HANDLE;
                MasterAxis := cam.AUX2;
                SlaveScaling := cam.F3;
            END_IF;
        ELSE
            Error := TRUE; ErrorID := cam.ERRID;
        END_IF;
    END_IF;
END_FUNCTION_BLOCK

(* ---- tc3_mc3ptp.st ---- *)
// Tc3_Mc3Ptp — MC3 point-to-point single-axis FBs missing from
// the Tc2_MC2 surface (TF55xx_MC3 bundle).
//
// Implemented over the builtin FB_MotionAxis (tplc-motion service):
//   MC_ReadActualTorque               torque actual (0x6077)
//   MC_ReadHardwareParameter          drive-param read (OD index)
//   MC_WriteHardwareParameter         drive-param write (OD index)
//   MC_WaitForStableActualPosition    velocity-window settle wait
//   MC_TriggerError                   fault inject (sim-ext 0x200D)
//   MC_SetHomingState                 accepted, no-op (documented)
//   MC_LoadControl                    accepted, no-op (documented)
//   MC_ActivateExternalSetpointGeneration  accepted, no-op
//
// Deviation notes: hardware parameters share the standard OD index
// space (TwinCAT drive-vendor parameter ids have no sim equivalent);
// SetHomingState/LoadControl/ActivateExternalSetpointGeneration
// configure drive-internal behaviour the simulated CiA402 drive does
// not model, so they complete with Done and change nothing; the
// camming (MC_Cam*), phasing (MC_Phasing*/MC_GearInPos/MC_HaltPhasing)
// and fluid-power (MC_ValveCharacterization) FBs plus the TcCOM
// AXIS_REF/ENCODER_AXIS_REF objects are deferred.

// ---- MC_ReadActualTorque: read actual torque (0x6077) ----
FUNCTION_BLOCK MC_ReadActualTorque
VAR_INPUT
    Enable : BOOL;
    Axis : UDINT;
END_VAR
VAR_OUTPUT
    Valid : BOOL;
    Torque : DINT;
    Busy : BOOL;
END_VAR
VAR
    ax : FB_MotionAxis;
END_VAR
    ax.OP := 3; ax();
    ax.AXIS := Axis;
    ax.OP := 4;
    ax.INDEX := 16#6077;
    ax();
    IF Enable AND ax.STATUS = 0 THEN
        Valid := TRUE;
        Torque := ax.VALUE;
    ELSE
        Valid := FALSE;
        Torque := 0;
    END_IF;
    Busy := FALSE;
END_FUNCTION_BLOCK

// ---- MC_ReadHardwareParameter: read a drive parameter ----
// ParameterNumber is the DS402 object-dictionary index, same
// convention as MC_ReadParameter.
FUNCTION_BLOCK MC_ReadHardwareParameter
VAR_INPUT
    Enable : BOOL;
    ParameterNumber : UDINT;
    Axis : UDINT;
END_VAR
VAR_OUTPUT
    Valid : BOOL;
    Value : DINT;
    Busy : BOOL;
END_VAR
VAR
    ax : FB_MotionAxis;
END_VAR
    ax.OP := 3; ax();
    ax.AXIS := Axis;
    ax.OP := 4;
    ax.INDEX := ParameterNumber;
    ax();
    IF Enable AND ax.STATUS = 0 THEN
        Valid := TRUE;
        Value := ax.VALUE;
    ELSE
        Valid := FALSE;
        Value := 0;
    END_IF;
    Busy := FALSE;
END_FUNCTION_BLOCK

// ---- MC_WriteHardwareParameter: write a drive parameter ----
FUNCTION_BLOCK MC_WriteHardwareParameter
VAR_INPUT
    Execute : BOOL;
    ParameterNumber : UDINT;
    Value : DINT;
    Axis : UDINT;
END_VAR
VAR_OUTPUT
    Done : BOOL;
    Busy : BOOL;
    Error : BOOL;
    ErrorID : UDINT;
END_VAR
VAR
    ax : FB_MotionAxis;
    exPrev : BOOL;
    exEdge : BOOL;
END_VAR
    ax.OP := 3; ax();
    ax.AXIS := Axis;
    exEdge := Execute AND NOT exPrev; exPrev := Execute;
    Done := FALSE; Error := FALSE; ErrorID := 0;
    IF exEdge THEN
        ax.OP := 5;
        ax.INDEX := ParameterNumber;
        ax.VALUE := Value;
        ax();
        IF ax.STATUS = 0 THEN
            Done := TRUE;
        ELSE
            Error := TRUE; ErrorID := ax.ERRID;
        END_IF;
    END_IF;
    Busy := FALSE;
END_FUNCTION_BLOCK

// ---- MC_WaitForStableActualPosition ----
// Execute edge arms the wait; Done fires once |VelocityActual|
// stays at or below VelocityWindow for SettleScans consecutive
// scans (position is implicitly stable because the sim integrates
// position from velocity). PositionWindow is accepted for
// signature fidelity: the sim exposes no sub-window position
// quantization, so only the velocity window gates completion.
FUNCTION_BLOCK MC_WaitForStableActualPosition
VAR_INPUT
    Execute : BOOL;
    PositionWindow : DINT;
    VelocityWindow : DINT;
    Axis : UDINT;
END_VAR
VAR_OUTPUT
    Done : BOOL;
    Busy : BOOL;
    Error : BOOL;
    ErrorID : UDINT;
END_VAR
VAR
    ax : FB_MotionAxis;
    exPrev : BOOL;
    exEdge : BOOL;
    armed : BOOL;
    still : INT;
    SettleScans : INT := 5;
END_VAR
    ax.AXIS := Axis;
    ax.OP := 3; ax();
    exEdge := Execute AND NOT exPrev; exPrev := Execute;
    Done := FALSE; Error := FALSE; ErrorID := 0;
    IF exEdge THEN
        armed := TRUE; still := 0;
    END_IF;
    IF armed THEN
        ax.OP := 6; ax();
        IF ax.STATUS < 0 THEN
            Error := TRUE; ErrorID := ax.ERRID; armed := FALSE;
        ELSIF ABS(ax.VEL_ACTUAL) <= VelocityWindow THEN
            still := still + 1;
            IF still >= SettleScans THEN
                Done := TRUE; armed := FALSE;
            END_IF;
        ELSE
            still := 0;
        END_IF;
    END_IF;
    Busy := armed;
END_FUNCTION_BLOCK

// ---- MC_TriggerError: inject a drive fault ----
// Writes ErrorCode to the sim-ext error-inject object (0x200D):
// nonzero latches the CiA402 fault state with that error code
// (readable via MC_ReadAxisError / 0x603F); write 0 to clear.
// ErrorCode 0 completes without faulting (used to clear).
FUNCTION_BLOCK MC_TriggerError
VAR_INPUT
    Execute : BOOL;
    ErrorCode : DINT;
    Axis : UDINT;
END_VAR
VAR_OUTPUT
    Done : BOOL;
    Busy : BOOL;
    Error : BOOL;
    ErrorID : UDINT;
END_VAR
VAR
    ax : FB_MotionAxis;
    exPrev : BOOL;
    exEdge : BOOL;
END_VAR
    ax.OP := 3; ax();
    ax.AXIS := Axis;
    exEdge := Execute AND NOT exPrev; exPrev := Execute;
    Done := FALSE; Error := FALSE; ErrorID := 0;
    IF exEdge THEN
        ax.OP := 5;
        ax.INDEX := 16#200D;
        ax.VALUE := ErrorCode;
        ax();
        IF ax.STATUS = 0 THEN
            Done := TRUE;
        ELSE
            Error := TRUE; ErrorID := ax.ERRID;
        END_IF;
    END_IF;
    Busy := FALSE;
END_FUNCTION_BLOCK

// ---- MC_SetHomingState: accepted no-op ----
// TwinCAT programs the drive homing state; the simulated drive
// derives homing state from the controlword, so the command
// completes with Done and HomingState is ignored.
FUNCTION_BLOCK MC_SetHomingState
VAR_INPUT
    Execute : BOOL;
    HomingState : UDINT;
    Axis : UDINT;
END_VAR
VAR_OUTPUT
    Done : BOOL;
    Busy : BOOL;
    Error : BOOL;
    ErrorID : UDINT;
END_VAR
VAR
    exPrev : BOOL;
    exEdge : BOOL;
END_VAR
    exEdge := Execute AND NOT exPrev; exPrev := Execute;
    Done := FALSE; Error := FALSE; ErrorID := 0;
    IF exEdge THEN Done := TRUE; END_IF;
    Busy := FALSE;
END_FUNCTION_BLOCK

// ---- MC_LoadControl: accepted no-op ----
// Loads controller parameters into the drive; the simulated drive
// has no separate control-parameter store, so the command
// completes with Done.
FUNCTION_BLOCK MC_LoadControl
VAR_INPUT
    Execute : BOOL;
    Axis : UDINT;
END_VAR
VAR_OUTPUT
    Done : BOOL;
    Busy : BOOL;
    Error : BOOL;
    ErrorID : UDINT;
END_VAR
VAR
    exPrev : BOOL;
    exEdge : BOOL;
END_VAR
    exEdge := Execute AND NOT exPrev; exPrev := Execute;
    Done := FALSE; Error := FALSE; ErrorID := 0;
    IF exEdge THEN Done := TRUE; END_IF;
    Busy := FALSE;
END_FUNCTION_BLOCK

// ---- MC_ActivateExternalSetpointGeneration: accepted no-op ----
// Selects drive-external setpoint generation; the sim has no
// external-setpoint mode distinct from the written targets, so the
// command completes with Done.
FUNCTION_BLOCK MC_ActivateExternalSetpointGeneration
VAR_INPUT
    Execute : BOOL;
    Axis : UDINT;
END_VAR
VAR_OUTPUT
    Done : BOOL;
    Busy : BOOL;
    Error : BOOL;
    ErrorID : UDINT;
END_VAR
VAR
    exPrev : BOOL;
    exEdge : BOOL;
END_VAR
    exEdge := Execute AND NOT exPrev; exPrev := Execute;
    Done := FALSE; Error := FALSE; ErrorID := 0;
    IF exEdge THEN Done := TRUE; END_IF;
    Busy := FALSE;
END_FUNCTION_BLOCK

(* ---- tc3_mcgroup.st ---- *)
// Tc3_McCoordinatedMotion — MC Group administration surface
// (TF5410 collision-avoidance / coordinated-motion bundle).
//
// This tranche implements the group bookkeeping FBs.  Motion
// execution (MC_MovePath, preparations, blockers, dwell), track
// following (MC_ActivateTrack, MC_TrackConveyorBelt,
// MC_ReadTrackPositions), collision-avoidance moves
// (MC_MoveAbsoluteCA etc.) and axis compensation
// (MC_RegisterCompensation, MC_TransformPosition) require the
// trajectory engine and are deferred.
//
// Flattened types (the ST dialect has no STRUCT/REFERENCE support):
//   AXES_GROUP_REF        -> AxesGroup : UDINT group handle (1..8)
//   AXIS_REF              -> Axis : UDINT axis handle
//   IDENT_IN_GROUP_REF    -> IdentInGroup : UDINT
//                            (UDINT_TO_IDENTINGROUP is the identity)
//   MC_COORD_REF          -> CoordTransform : UDINT
//   ECmSetpointSource     -> SetpointSource : UDINT
//                            (1=Group, 2=MCS, 3=ACS)
//   MC_LREAL              -> LREAL
//
// Group states (approximation of TwinCAT mcGroupState*):
//   0 empty, 1 disabled, 2 standby, 3 moving, 4 error-disabled,
//   5 group-error.  The service is synchronous, so Busy stays
//   FALSE and Done/Error pulse on the execute scan.
//   ErrorId carries the service status magnitude.

// ---- UDINT_TO_IDENTINGROUP: identity conversion ----
FUNCTION UDINT_TO_IDENTINGROUP : UDINT
VAR_INPUT
    InVal : UDINT;
END_VAR
UDINT_TO_IDENTINGROUP := InVal;
END_FUNCTION

// ---- shared command skeleton: rising-edge Execute -> FB_McGroup --
// Each public FB owns one FB_McGroup instance `mg`.

FUNCTION_BLOCK MC_AddAxisToGroup
VAR_INPUT
    Execute : BOOL;
    IdentInGroup : UDINT;
END_VAR
VAR_IN_OUT
    AxesGroup : UDINT;
    Axis : UDINT;
END_VAR
VAR_OUTPUT
    Done : BOOL;
    Busy : BOOL;
    Error : BOOL;
    ErrorId : UDINT;
END_VAR
VAR
    mg : FB_McGroup;
    exPrev : BOOL;
    edge : BOOL;
    ok : BOOL;
END_VAR
ok := FALSE;
edge := Execute AND NOT exPrev;
IF edge THEN
    mg.OP := 1; mg.GRP := AxesGroup; mg();
    AxesGroup := mg.GRP;
    mg.OP := 2; mg.AXIS := Axis; mg.IDENT := IdentInGroup; mg();
    IF mg.STATUS = 0 THEN ok := TRUE; END_IF;
END_IF;
exPrev := Execute;
Done := ok; Busy := FALSE;
Error := edge AND NOT ok AND mg.STATUS <> 0;
IF edge AND mg.STATUS < 0 THEN ErrorId := 0 - mg.STATUS; END_IF;
END_FUNCTION_BLOCK

FUNCTION_BLOCK MC_RemoveAxisFromGroup
VAR_INPUT
    Execute : BOOL;
    IdentInGroup : UDINT;
END_VAR
VAR_IN_OUT
    AxesGroup : UDINT;
    Axis : UDINT;
END_VAR
VAR_OUTPUT
    Done : BOOL;
    Busy : BOOL;
    Error : BOOL;
    ErrorId : UDINT;
END_VAR
VAR
    mg : FB_McGroup;
    exPrev : BOOL;
    edge : BOOL;
    ok : BOOL;
END_VAR
ok := FALSE;
edge := Execute AND NOT exPrev;
IF edge THEN
    mg.OP := 1; mg.GRP := AxesGroup; mg();
    AxesGroup := mg.GRP;
    mg.OP := 3; mg.AXIS := Axis; mg.IDENT := IdentInGroup; mg();
    IF mg.STATUS = 0 THEN ok := TRUE; END_IF;
END_IF;
exPrev := Execute;
Done := ok; Busy := FALSE;
Error := edge AND NOT ok AND mg.STATUS <> 0;
IF edge AND mg.STATUS < 0 THEN ErrorId := 0 - mg.STATUS; END_IF;
END_FUNCTION_BLOCK

FUNCTION_BLOCK MC_UngroupAllAxes
VAR_INPUT
    Execute : BOOL;
END_VAR
VAR_IN_OUT
    AxesGroup : UDINT;
END_VAR
VAR_OUTPUT
    Done : BOOL;
    Busy : BOOL;
    Error : BOOL;
    ErrorId : UDINT;
END_VAR
VAR
    mg : FB_McGroup;
    exPrev : BOOL;
    edge : BOOL;
    ok : BOOL;
END_VAR
ok := FALSE;
edge := Execute AND NOT exPrev;
IF edge THEN
    mg.OP := 4; mg.GRP := AxesGroup; mg();
    IF mg.STATUS = 0 THEN ok := TRUE; END_IF;
END_IF;
exPrev := Execute;
Done := ok; Busy := FALSE;
Error := edge AND NOT ok AND mg.STATUS <> 0;
IF edge AND mg.STATUS < 0 THEN ErrorId := 0 - mg.STATUS; END_IF;
END_FUNCTION_BLOCK

FUNCTION_BLOCK MC_GroupEnable
VAR_INPUT
    Execute : BOOL;
END_VAR
VAR_IN_OUT
    AxesGroup : UDINT;
END_VAR
VAR_OUTPUT
    Done : BOOL;
    Busy : BOOL;
    Error : BOOL;
    ErrorId : UDINT;
END_VAR
VAR
    mg : FB_McGroup;
    exPrev : BOOL;
    edge : BOOL;
    ok : BOOL;
END_VAR
ok := FALSE;
edge := Execute AND NOT exPrev;
IF edge THEN
    mg.OP := 1; mg.GRP := AxesGroup; mg();
    AxesGroup := mg.GRP;
    mg.OP := 5; mg.ENABLE := 1; mg();
    IF mg.STATUS = 0 THEN ok := TRUE; END_IF;
END_IF;
exPrev := Execute;
Done := ok; Busy := FALSE;
Error := edge AND NOT ok AND mg.STATUS <> 0;
IF edge AND mg.STATUS < 0 THEN ErrorId := 0 - mg.STATUS; END_IF;
END_FUNCTION_BLOCK

FUNCTION_BLOCK MC_GroupDisable
VAR_INPUT
    Execute : BOOL;
END_VAR
VAR_IN_OUT
    AxesGroup : UDINT;
END_VAR
VAR_OUTPUT
    Done : BOOL;
    Busy : BOOL;
    Error : BOOL;
    ErrorId : UDINT;
END_VAR
VAR
    mg : FB_McGroup;
    exPrev : BOOL;
    edge : BOOL;
    ok : BOOL;
END_VAR
ok := FALSE;
edge := Execute AND NOT exPrev;
IF edge THEN
    mg.OP := 1; mg.GRP := AxesGroup; mg();
    AxesGroup := mg.GRP;
    mg.OP := 5; mg.ENABLE := 0; mg();
    IF mg.STATUS = 0 THEN ok := TRUE; END_IF;
END_IF;
exPrev := Execute;
Done := ok; Busy := FALSE;
Error := edge AND NOT ok AND mg.STATUS <> 0;
IF edge AND mg.STATUS < 0 THEN ErrorId := 0 - mg.STATUS; END_IF;
END_FUNCTION_BLOCK

FUNCTION_BLOCK MC_GroupReset
VAR_INPUT
    Execute : BOOL;
END_VAR
VAR_IN_OUT
    AxesGroup : UDINT;
END_VAR
VAR_OUTPUT
    Done : BOOL;
    Busy : BOOL;
    Error : BOOL;
    ErrorId : UDINT;
END_VAR
VAR
    mg : FB_McGroup;
    exPrev : BOOL;
    edge : BOOL;
    ok : BOOL;
END_VAR
ok := FALSE;
edge := Execute AND NOT exPrev;
IF edge THEN
    mg.OP := 1; mg.GRP := AxesGroup; mg();
    AxesGroup := mg.GRP;
    mg.OP := 5; mg.ENABLE := 2; mg();
    IF mg.STATUS = 0 THEN ok := TRUE; END_IF;
END_IF;
exPrev := Execute;
Done := ok; Busy := FALSE;
Error := edge AND NOT ok AND mg.STATUS <> 0;
IF edge AND mg.STATUS < 0 THEN ErrorId := 0 - mg.STATUS; END_IF;
END_FUNCTION_BLOCK

// ---- level-triggered status readers (Enable input) ----

FUNCTION_BLOCK MC_GroupReadStatus
VAR_INPUT
    Enable : BOOL;
END_VAR
VAR_IN_OUT
    AxesGroup : UDINT;
END_VAR
VAR_OUTPUT
    Valid : BOOL;
    Busy : BOOL;
    GroupMoving : BOOL;
    GroupHoming : BOOL;
    GroupErrorStop : BOOL;
    GroupNotReady : BOOL;
    GroupStandby : BOOL;
    GroupStopping : BOOL;
    GroupDisabled : BOOL;
    AllAxesStanding : BOOL;
    InPosition : BOOL;
    Error : BOOL;
    ErrorId : UDINT;
END_VAR
VAR
    mg : FB_McGroup;
END_VAR
Valid := FALSE; Busy := FALSE; Error := FALSE; ErrorId := 0;
GroupMoving := FALSE; GroupHoming := FALSE; GroupErrorStop := FALSE;
GroupNotReady := FALSE; GroupStandby := FALSE; GroupStopping := FALSE;
GroupDisabled := FALSE; AllAxesStanding := FALSE; InPosition := FALSE;
IF Enable THEN
    mg.OP := 6; mg.GRP := AxesGroup; mg();
    IF mg.STATUS = 0 THEN
        Valid := TRUE;
        GroupMoving := mg.STATE = 3;
        GroupStandby := mg.STATE = 2;
        GroupDisabled := mg.STATE = 0 OR mg.STATE = 1 OR
                        mg.STATE = 4;
        AllAxesStanding := mg.STATE = 2 OR mg.STATE = 3;
        /* GroupHoming/GroupErrorStop/GroupNotReady/GroupStopping/
           InPosition need the motion engine; always FALSE here. */
    ELSE
        Error := TRUE;
        IF mg.STATUS < 0 THEN ErrorId := (0 - mg.STATUS); END_IF;
    END_IF;
END_IF;
END_FUNCTION_BLOCK

FUNCTION_BLOCK MC_GroupReadError
VAR_INPUT
    Enable : BOOL;
END_VAR
VAR_IN_OUT
    AxesGroup : UDINT;
END_VAR
VAR_OUTPUT
    Valid : BOOL;
    Busy : BOOL;
    Error : BOOL;
    ErrorId : UDINT;
    GroupErrorId : UDINT;
END_VAR
VAR
    mg : FB_McGroup;
END_VAR
Valid := FALSE; Busy := FALSE; Error := FALSE;
ErrorId := 0; GroupErrorId := 0;
IF Enable THEN
    mg.OP := 6; mg.GRP := AxesGroup; mg();
    IF mg.STATUS = 0 THEN
        Valid := TRUE;
        GroupErrorId := mg.ERRID;
    ELSE
        Error := TRUE;
        IF mg.STATUS < 0 THEN ErrorId := (0 - mg.STATUS); END_IF;
    END_IF;
END_IF;
END_FUNCTION_BLOCK

FUNCTION_BLOCK MC_GroupSetOverride
VAR_INPUT
    Execute : BOOL;
    Enable : BOOL;
    VelFactor : LREAL;
END_VAR
VAR_IN_OUT
    AxesGroup : UDINT;
END_VAR
VAR_OUTPUT
    Done : BOOL;
    Busy : BOOL;
    Error : BOOL;
    ErrorId : UDINT;
    OverrideActual : LREAL;
END_VAR
VAR
    mg : FB_McGroup;
    exPrev : BOOL;
    edge : BOOL;
    ok : BOOL;
    ovr : LREAL;
END_VAR
ok := FALSE; ovr := 1.0;
edge := Execute AND NOT exPrev;
IF Enable THEN ovr := VelFactor; END_IF;
IF edge THEN
    mg.OP := 1; mg.GRP := AxesGroup; mg();
    AxesGroup := mg.GRP;
    mg.OP := 7; mg.OVR := ovr; mg();
    IF mg.STATUS = 0 THEN
        ok := TRUE;
        OverrideActual := mg.OVRACT;
    END_IF;
END_IF;
exPrev := Execute;
Done := ok; Busy := FALSE;
Error := edge AND NOT ok AND mg.STATUS <> 0;
IF edge AND mg.STATUS < 0 THEN ErrorId := 0 - mg.STATUS; END_IF;
END_FUNCTION_BLOCK

FUNCTION_BLOCK MC_GroupSetSetpointSource
VAR_INPUT
    Execute : BOOL;
    SetpointSource : UDINT;
END_VAR
VAR_IN_OUT
    AxesGroup : UDINT;
END_VAR
VAR_OUTPUT
    Done : BOOL;
    Busy : BOOL;
    Error : BOOL;
    ErrorId : UDINT;
END_VAR
VAR
    mg : FB_McGroup;
    exPrev : BOOL;
    edge : BOOL;
    ok : BOOL;
    src : UDINT;
END_VAR
ok := FALSE;
edge := Execute AND NOT exPrev;
src := SetpointSource - 1; /* 1/2/3 -> 0/1/2 */
IF edge THEN
    mg.OP := 1; mg.GRP := AxesGroup; mg();
    AxesGroup := mg.GRP;
    mg.OP := 8; mg.SOURCE := src; mg();
    IF mg.STATUS = 0 THEN ok := TRUE; END_IF;
END_IF;
exPrev := Execute;
Done := ok; Busy := FALSE;
Error := edge AND NOT ok AND mg.STATUS <> 0;
IF edge AND mg.STATUS < 0 THEN ErrorId := 0 - mg.STATUS; END_IF;
END_FUNCTION_BLOCK

FUNCTION_BLOCK MC_SetCoordinateTransform
VAR_INPUT
    Execute : BOOL;
    CoordTransform : UDINT;
END_VAR
VAR_IN_OUT
    AxesGroup : UDINT;
END_VAR
VAR_OUTPUT
    Done : BOOL;
    Busy : BOOL;
    Active : BOOL;
    CommandAborted : BOOL;
    Error : BOOL;
    ErrorId : UDINT;
END_VAR
VAR
    mg : FB_McGroup;
    exPrev : BOOL;
    edge : BOOL;
    ok : BOOL;
    act : BOOL;
END_VAR
ok := FALSE;
edge := Execute AND NOT exPrev;
IF edge THEN
    mg.OP := 1; mg.GRP := AxesGroup; mg();
    AxesGroup := mg.GRP;
    mg.OP := 9; mg.COORD := CoordTransform; mg();
    IF mg.STATUS = 0 THEN ok := TRUE; act := TRUE; END_IF;
END_IF;
exPrev := Execute;
Done := ok; Busy := FALSE; CommandAborted := FALSE;
Active := act;
Error := edge AND NOT ok AND mg.STATUS <> 0;
IF edge AND mg.STATUS < 0 THEN ErrorId := 0 - mg.STATUS; END_IF;
END_FUNCTION_BLOCK

// ---- MC_GroupStop / MC_GroupHalt: stop every axis in the group ----
// The group membership lives in tplc-mcgroup; the per-axis stop is
// applied through FB_MotionAxis. MC_GroupStop ramps each axis to
// rest in PV mode (0x60FF=0, the decelerated-stop shape); its
// Deceleration input is accepted but the simulated drive applies
// its own ramp. MC_GroupHalt disables each axis immediately
// (controlword 0x000B). Both poll VEL_ACTUAL and report Done once
// every member reads zero velocity.

FUNCTION_BLOCK MC_GroupStop
VAR_INPUT
    Execute : BOOL;
    Deceleration : LREAL := 0.0;
END_VAR
VAR_IN_OUT
    AxesGroup : UDINT;
END_VAR
VAR_OUTPUT
    Done : BOOL;
    Busy : BOOL;
    Error : BOOL;
    ErrorId : UDINT;
END_VAR
VAR
    mg : FB_McGroup;
    ax : FB_MotionAxis;
    exPrev : BOOL;
    exEdge : BOOL;
    active : BOOL;
    issued : BOOL;
    i : UDINT;
    n : UDINT;
    stopped : UDINT;
    axh : UDINT;
END_VAR
    mg.GRP := AxesGroup;
    mg.OP := 10; mg();
    AxesGroup := mg.GRP;
    n := mg.NAXES;
    exEdge := Execute AND NOT exPrev; exPrev := Execute;
    Done := FALSE; Busy := FALSE;
    Error := FALSE; ErrorId := 0;
    IF exEdge THEN active := TRUE; issued := FALSE; END_IF;
    IF active THEN
        IF NOT issued THEN
            FOR i := 0 TO 15 DO
                IF i < n THEN
                    axh := mg.AXES[i];
                    ax.AXIS := axh;
                    ax.OP := 5; ax.INDEX := 16#6040; ax.VALUE := 16#000F; ax();
                    ax.OP := 5; ax.INDEX := 16#6060; ax.VALUE := 3; ax();
                    ax.OP := 5; ax.INDEX := 16#60FF; ax.VALUE := 0; ax();
                END_IF;
            END_FOR;
            issued := TRUE;
        END_IF;
        stopped := 0;
        FOR i := 0 TO 15 DO
            IF i < n THEN
                axh := mg.AXES[i];
                ax.AXIS := axh; ax.OP := 3; ax();
                ax.OP := 6; ax();
                IF ax.VEL_ACTUAL = 0 THEN stopped := stopped + 1; END_IF;
            END_IF;
        END_FOR;
        IF n = 0 OR stopped >= n THEN
            Done := TRUE; active := FALSE;
        END_IF;
        Busy := active;
        IF mg.STATUS < 0 THEN
            Error := TRUE; ErrorId := 0 - mg.STATUS; active := FALSE;
        END_IF;
    END_IF;
END_FUNCTION_BLOCK

FUNCTION_BLOCK MC_GroupHalt
VAR_INPUT
    Execute : BOOL;
END_VAR
VAR_IN_OUT
    AxesGroup : UDINT;
END_VAR
VAR_OUTPUT
    Done : BOOL;
    Busy : BOOL;
    Error : BOOL;
    ErrorId : UDINT;
END_VAR
VAR
    mg : FB_McGroup;
    ax : FB_MotionAxis;
    exPrev : BOOL;
    exEdge : BOOL;
    active : BOOL;
    issued : BOOL;
    i : UDINT;
    n : UDINT;
    stopped : UDINT;
    axh : UDINT;
END_VAR
    mg.GRP := AxesGroup;
    mg.OP := 10; mg();
    AxesGroup := mg.GRP;
    n := mg.NAXES;
    exEdge := Execute AND NOT exPrev; exPrev := Execute;
    Done := FALSE; Busy := FALSE;
    Error := FALSE; ErrorId := 0;
    IF exEdge THEN active := TRUE; issued := FALSE; END_IF;
    IF active THEN
        IF NOT issued THEN
            FOR i := 0 TO 15 DO
                IF i < n THEN
                    axh := mg.AXES[i];
                    ax.AXIS := axh;
                    ax.OP := 5; ax.INDEX := 16#6040; ax.VALUE := 16#000B; ax();
                END_IF;
            END_FOR;
            issued := TRUE;
        END_IF;
        stopped := 0;
        FOR i := 0 TO 15 DO
            IF i < n THEN
                axh := mg.AXES[i];
                ax.AXIS := axh; ax.OP := 3; ax();
                ax.OP := 6; ax();
                IF ax.VEL_ACTUAL = 0 THEN stopped := stopped + 1; END_IF;
            END_IF;
        END_FOR;
        IF n = 0 OR stopped >= n THEN
            Done := TRUE; active := FALSE;
        END_IF;
        Busy := active;
        IF mg.STATUS < 0 THEN
            Error := TRUE; ErrorId := 0 - mg.STATUS; active := FALSE;
        END_IF;
    END_IF;
END_FUNCTION_BLOCK
